{region 'Documentation'}
(*!
<summary>Restarts the scenario sequence and outer checks.</summary>
*)
{endregion}
METHOD PROTECTED ProcessReset
FScenario := ScenarioLowerLimits;
FChecked := FALSE;
FSubjectEnable := FALSE;
FEvaluateSubjects := FALSE;
FObservationReady := FALSE;
FFirstFailedScenario := 0;
FFailedDuringEvaluation := FALSE;
FCapture.Reset();
ResetSubjects();
FResults.Reset();
FActivity.Reset();
FInputs.Reset();
FFindings.Reset();
CompleteReset();
END_METHOD

{region 'Documentation'}
(*!
<summary>Consumes reset, evaluates, then waits for the outer checks before advancing.</summary>
*)
{endregion}
METHOD PROTECTED ProcessTests
VAR_INPUT
    Enable : BOOL; //! Phase permission supplied by the owning Test Case; FALSE does not authorize progression, while observation may continue.
END_VAR
IF NOT Enable THEN
    RETURN;
END_IF;

IF FChecked THEN
    FChecked := FALSE;
    FObservationReady := FALSE;
    IF FEvaluateSubjects THEN
        IF FScenario = LastScenario THEN
            CompleteTests();
            RETURN;
        END_IF;
        FScenario := FScenario + 1;
    END_IF;
    FEvaluateSubjects := NOT FEvaluateSubjects;
END_IF;

IF NOT SelectScenario() THEN
    RETURN;
END_IF;
FCapture.Reset();
IF NOT FEvaluateSubjects THEN
    ResetSubjects();
END_IF;

CallSubjects();
CheckResults();
CheckInputs();
CheckFindings();
IF (FFirstFailedScenario = 0)
    AND NOT (FResultsMatch AND FActivityMatch AND FInputsMatch AND FFindingsMatch) THEN
    FFirstFailedScenario := FScenario;
    FFailedDuringEvaluation := FEvaluateSubjects;
END_IF;
FObservationReady := TRUE;
END_METHOD

{region 'Documentation'}
(*!
<summary>Queues reset; the next bound FB call consumes it without evaluating.</summary>
*)
{endregion}
METHOD PRIVATE ResetSubjects
FSigned.Reset();
FUnsigned.Reset();
END_METHOD

{region 'Documentation'}
(*!
<summary>Selects explicit stimuli and expected results for one scenario.</summary>
*)
{endregion}
METHOD PRIVATE SelectScenario : BOOL //! TRUE after selecting a supported scenario and its literal expectations; FALSE reports an unknown scenario.
SelectScenario := FALSE;
FSubjectEnable := TRUE;
FSignedValue := -127;
FSignedMinimum := -128;
FUnsignedValue := 128;
FUnsignedMinimum := 128;
FUnsignedMaximum := 255;
CASE FScenario OF
    ScenarioLowerLimits:
        FSignedExpectedResult := E_Result.Passed;
        FSignedExpectedFinding := FALSE;
        FUnsignedExpectedResult := E_Result.Passed;
        FUnsignedExpectedFinding := FALSE;
    ScenarioUpperLimits:
        FSignedValue := 127;
        FUnsignedValue := 255;
        FSignedExpectedResult := E_Result.Passed;
        FSignedExpectedFinding := FALSE;
        FUnsignedExpectedResult := E_Result.Passed;
        FUnsignedExpectedFinding := FALSE;
    ScenarioEqualSignedMinimum:
        FSignedValue := -128;
        FSignedExpectedResult := E_Result.Failed;
        FSignedExpectedFinding := TRUE;
        FUnsignedExpectedResult := E_Result.Passed;
        FUnsignedExpectedFinding := FALSE;
    ScenarioOutsideRange:
        FSignedValue := -128;
        FSignedMinimum := -127;
        FUnsignedValue := 127;
        FSignedExpectedResult := E_Result.Failed;
        FSignedExpectedFinding := TRUE;
        FUnsignedExpectedResult := E_Result.Failed;
        FUnsignedExpectedFinding := TRUE;
    ScenarioAboveMaximum:
        FUnsignedValue := 255;
        FUnsignedMaximum := 254;
        FSignedExpectedResult := E_Result.Passed;
        FSignedExpectedFinding := FALSE;
        FUnsignedExpectedResult := E_Result.Failed;
        FUnsignedExpectedFinding := TRUE;
    ScenarioSingleValue:
        FUnsignedMinimum := 255;
        FUnsignedMaximum := 255;
        FUnsignedValue := 255;
        FSignedExpectedResult := E_Result.Passed;
        FSignedExpectedFinding := FALSE;
        FUnsignedExpectedResult := E_Result.Passed;
        FUnsignedExpectedFinding := FALSE;
    ScenarioReversedRange:
        FUnsignedMinimum := 255;
        FUnsignedMaximum := 128;
        FSignedExpectedResult := E_Result.Passed;
        FSignedExpectedFinding := FALSE;
        FUnsignedExpectedResult := E_Result.Error;
        FUnsignedExpectedFinding := TRUE;
ELSE
    Error(Message := 'Unknown variant Assertion scenario.');
    RETURN;
END_CASE;

SelectScenario := TRUE;
END_METHOD

END_FUNCTION_BLOCK

// ---- SelfTests/TestCases/TestSuite_AssertionVariants/Test_AssertionTemporalVariants.TcPOU
{region 'Documentation'}
(*!
<summary>Checks temporal variants with isolated production subjects.</summary>
<description>
Each independent scenario consumes a bound reset call before its evaluation call.
ProcessAssertions checks the observation before ProcessTests advances.
SelectScenario holds explicit expected results; no production algorithm is mirrored.
Expected findings remain in the local capture; only outer checks affect the test result.
FirstFailedScenario and FailedDuringEvaluation retain the first mismatch.
Each scenario uses literal typed inputs at the declared operand widths.
</description>
*)
{endregion}
FUNCTION_BLOCK Test_AssertionTemporalVariants EXTENDS TestCaseBase
VAR
    FTimestamp : AssertEqual_LDT;
    FTimestampExpectedResult : E_Result;
    FTimestampExpectedFinding : BOOL;
    FTimespan : AssertInTimespan_DT;
    FTimespanExpectedResult : E_Result;
    FTimespanExpectedFinding : BOOL;

    FTimestampValue : LDT;
    FExpectedTimestamp : LDT;
    FTime : DT;
    FStartTime : DT;
    FEndTime : DT;
    FSubjectEnable : BOOL;
    FCapture : EventBuffer;
    FEvents : ARRAY[1..CaptureLength] OF ST_Event;
    FCaptureFifo : ST_FifoStatus;
    FCaptureStatus : ST_EventBufferStatus;
    FSetupValid : BOOL;
    FScenario : UINT;
    FChecked : BOOL;
    FEvaluateSubjects : BOOL;
    FObservationReady : BOOL;
    FFirstFailedScenario : UINT;
    FFailedDuringEvaluation : BOOL;
    FResultsMatch : BOOL;
    FResults : AssertTrue;
    FActivityMatch : BOOL;
    FActivity : AssertTrue;
    FInputsMatch : BOOL;
    FInputs : AssertTrue;
    FFindingsMatch : BOOL;
    FFindings : AssertTrue;
END_VAR
VAR CONSTANT
    CaptureLength : UINT := 8;
    ScenarioLowerBound : UINT := 1;
    ScenarioUpperBound : UINT := 2;
    ScenarioNanosecondDifference : UINT := 3;
    ScenarioBeforeStart : UINT := 4;
    ScenarioAfterEnd : UINT := 5;
    ScenarioSingleInstant : UINT := 6;
    ScenarioReversedTimespan : UINT := 7;
    LastScenario : UINT := ScenarioReversedTimespan;
END_VAR

SUPER^();

{region 'Documentation'}
(*!
<summary>Aggregates only outer checks, not intentionally failing subjects.</summary>
*)
{endregion}
METHOD PROTECTED AggregateResults
VAR_INPUT
    Aggregator : I_ResultAggregator; //! Borrowed result sink owned by the outer Test Case; add this test's checking Assertions without resetting or retaining the sink.
END_VAR
Aggregator.AddProvider(Provider := FResults);
Aggregator.AddProvider(Provider := FActivity);
Aggregator.AddProvider(Provider := FInputs);
Aggregator.AddProvider(Provider := FFindings);
END_METHOD

{region 'Documentation'}
(*!
<summary>Calls each inherited production subject once with caller-owned input storage.</summary>
*)
{endregion}
METHOD PRIVATE CallSubjects
FTimestamp(Enable := FSubjectEnable,
    State := E_State.Running,
    IN := FTimestampValue,
    Expected := FExpectedTimestamp);
FTimespan(Enable := FSubjectEnable,
    State := E_State.Running,
    IN := FTime,
    StartTime := FStartTime,
    EndTime := FEndTime);
END_METHOD

{region 'Documentation'}
(*!
<summary>Checks one subject finding in call order; expected outcomes come from the scenario.</summary>
*)
{endregion}
METHOD PRIVATE CheckFinding : BOOL //! TRUE when the required finding checks pass; calls requiring no finding also succeed.
VAR_INPUT
    Subject : I_Assertion; //! Assertion interface supplying the expected finding identity.
    ExpectedResult : E_Result; //! Independently authored result expected in the captured finding.
    ExpectedFinding : BOOL; //! TRUE when this scenario requires a finding during active evaluation.
END_VAR
VAR_IN_OUT
    Index : UINT; //! One-based next finding index; advanced when this call checks a required finding.
END_VAR
CheckFinding := TRUE;
IF FEvaluateSubjects AND ExpectedFinding THEN
    CheckFinding := (FEvents[Index].SequenceId = UINT_TO_UDINT(Index))
        AND (FEvents[Index].Name = Subject.Name)
        AND (FEvents[Index].OwnerScope = E_OwnerScope.Assertion)
        AND (FEvents[Index].EventType = E_EventType.Result)
        AND (FEvents[Index].State = E_State.Running)
        AND (FEvents[Index].Result = ExpectedResult)
        AND (FEvents[Index].Message <> '');
    Index := Index + 1;
END_IF;
END_METHOD

{region 'Documentation'}
(*!
<summary>Checks exact finding count and identities; at most one finding per subject.</summary>
*)
{endregion}
METHOD PRIVATE CheckFindings
VAR
    Index : UINT;
    Matches : BOOL;
END_VAR
Index := 1;
FFindingsMatch := TRUE;
Matches := CheckFinding(Subject := FTimestamp,
    ExpectedResult := FTimestampExpectedResult,
    ExpectedFinding := FTimestampExpectedFinding,
    Index := Index);
FFindingsMatch := FFindingsMatch AND Matches;
Matches := CheckFinding(Subject := FTimespan,
    ExpectedResult := FTimespanExpectedResult,
    ExpectedFinding := FTimespanExpectedFinding,
    Index := Index);
FFindingsMatch := FFindingsMatch AND Matches;
FFindingsMatch := FFindingsMatch
    AND (FCaptureStatus.SequenceId = UINT_TO_UDINT(Index - 1))
    AND (FCaptureStatus.LostEventCount = 0);
END_METHOD

{region 'Documentation'}
(*!
<summary>Rejects incomplete subject, capture or outer Assertion setup.</summary>
*)
{endregion}
METHOD PROTECTED CheckInitialization : BOOL //! TRUE when the inherited initialization check and this concrete fixture check both accept the setup.
CheckInitialization := SUPER^.CheckInitialization();
IF NOT CheckInitialization THEN
    RETURN;
END_IF;

CheckInitialization := FSetupValid
    AND FResults.IsInitialized
    AND FActivity.IsInitialized
    AND FInputs.IsInitialized
    AND FFindings.IsInitialized;
IF NOT CheckInitialization THEN
    EventPublisher.PublishEvent(Event := CreateFrameworkEvent(Name := Name,
        ResourceName := '',
        State := State,
        Severity := E_EventSeverity.Error,
        Message := 'Variant selftest setup failed.'));
END_IF;
END_METHOD

{region 'Documentation'}
(*!
<summary>Verifies input preservation without using the tested comparison algorithm.</summary>
*)
{endregion}
METHOD PRIVATE CheckInputs
FInputsMatch := (FTimestamp.IN = FTimestampValue)
    AND (FTimestamp.Expected = FExpectedTimestamp)
    AND (FTimespan.IN = FTime)
    AND (FTimespan.StartTime = FStartTime)
    AND (FTimespan.EndTime = FEndTime);
END_METHOD

{region 'Documentation'}
(*!
<summary>Checks literal evaluation results, or NotEvaluated on the reset call.</summary>
*)
{endregion}
METHOD PRIVATE CheckResults
IF FEvaluateSubjects THEN
    FResultsMatch := (FTimestamp.Result = FTimestampExpectedResult)
        AND (FTimespan.Result = FTimespanExpectedResult);
ELSE
    FResultsMatch := (FTimestamp.Result = E_Result.NotEvaluated)
        AND (FTimespan.Result = E_Result.NotEvaluated);
END_IF;
FActivityMatch := (FTimestamp.Enabled = FSubjectEnable)
    AND (FTimestamp.ObservationActive = (FEvaluateSubjects AND FSubjectEnable))
    AND (FTimestamp.EvaluationActive = (FEvaluateSubjects AND FSubjectEnable))
    AND (FTimespan.Enabled = FSubjectEnable)
    AND (FTimespan.ObservationActive = (FEvaluateSubjects AND FSubjectEnable))
    AND (FTimespan.EvaluationActive = (FEvaluateSubjects AND FSubjectEnable));
END_METHOD

{region 'Documentation'}
(*!
<summary>Initializes outer checks and isolates intentional subject findings.</summary>
*)
{endregion}
METHOD PROTECTED Configure
VAR
    Initialized : BOOL;
END_VAR
FPreparationStateCount := 0;
FTestStateCount := 1;
FResults.Initialize(Parent := THIS^,
    AssertionName := 'Results');
FActivity.Initialize(Parent := THIS^,
    AssertionName := 'Activity');
FInputs.Initialize(Parent := THIS^,
    AssertionName := 'Inputs');
FFindings.Initialize(Parent := THIS^,
    AssertionName := 'Findings');
FSetupValid := FCapture.Initialize(Buffer := FEvents,
    FifoControl := FCaptureFifo,
    Status := FCaptureStatus);
FTimestamp.BindPublisher(Publisher := FCapture);
Initialized := FTimestamp.Initialize(Parent := THIS^,
    AssertionName := 'Timestamp');
FSetupValid := FSetupValid AND Initialized;
FTimespan.BindPublisher(Publisher := FCapture);
Initialized := FTimespan.Initialize(Parent := THIS^,
    AssertionName := 'Timespan');
FSetupValid := FSetupValid AND Initialized;
END_METHOD

{region 'Documentation'}
(*!
<summary>Completes abort; no asynchronous resource is owned.</summary>
*)
{endregion}
METHOD PROTECTED ProcessAbort
VAR_INPUT
    Enable : BOOL; //! Phase permission supplied by the owning Test Case; FALSE does not authorize progression, while observation may continue.
END_VAR
IF Enable THEN
    CompleteAbort();
END_IF;
END_METHOD

{region 'Documentation'}
(*!
<summary>Latches this call's checks before progression is permitted.</summary>
*)
{endregion}
METHOD PROTECTED ProcessAssertions
VAR_INPUT
    Enable : BOOL; //! Phase permission supplied by the owning Test Case; FALSE does not authorize progression, while observation may continue.
END_VAR
VAR
    Check : BOOL;
END_VAR
Check := Enable AND FObservationReady;
FResults(Enable := Check,
    State := State,
    IN := FResultsMatch);
FActivity(Enable := Check,
    State := State,
    IN := FActivityMatch);
FInputs(Enable := Check,
    State := State,
    IN := FInputsMatch);
FFindings(Enable := Check,
    State := State,
    IN := FFindingsMatch);
IF Check THEN
    FChecked := TRUE;
END_IF;
END_METHOD

{region 'Documentation'}
(*!
<summary>No Preparation phase is needed.</summary>
*)
{endregion}
METHOD PROTECTED ProcessPreparations
VAR_INPUT
    // SA0033: Required hook; this test has no Preparation phase.
    {attribute 'analysis' := '-33'}
    Enable : BOOL; //! Phase permission supplied by the owning Test Case; FALSE does not authorize progression, while observation may continue.
END_VAR
END_METHOD

{region 'Documentation'}
(*!
<summary>Restarts the scenario sequence and outer checks.</summary>
*)
{endregion}
METHOD PROTECTED ProcessReset
FScenario := ScenarioLowerBound;
FChecked := FALSE;
FSubjectEnable := FALSE;
FEvaluateSubjects := FALSE;
FObservationReady := FALSE;
FFirstFailedScenario := 0;
FFailedDuringEvaluation := FALSE;
FCapture.Reset();
ResetSubjects();
FResults.Reset();
FActivity.Reset();
FInputs.Reset();
FFindings.Reset();
CompleteReset();
END_METHOD

{region 'Documentation'}
(*!
<summary>Consumes reset, evaluates, then waits for the outer checks before advancing.</summary>
*)
{endregion}
METHOD PROTECTED ProcessTests
VAR_INPUT
    Enable : BOOL; //! Phase permission supplied by the owning Test Case; FALSE does not authorize progression, while observation may continue.
END_VAR
IF NOT Enable THEN
    RETURN;
END_IF;

IF FChecked THEN
    FChecked := FALSE;
    FObservationReady := FALSE;
    IF FEvaluateSubjects THEN
        IF FScenario = LastScenario THEN
            CompleteTests();
            RETURN;
        END_IF;
        FScenario := FScenario + 1;
    END_IF;
    FEvaluateSubjects := NOT FEvaluateSubjects;
END_IF;

IF NOT SelectScenario() THEN
    RETURN;
END_IF;
FCapture.Reset();
IF NOT FEvaluateSubjects THEN
    ResetSubjects();
END_IF;

CallSubjects();
CheckResults();
CheckInputs();
CheckFindings();
IF (FFirstFailedScenario = 0)
    AND NOT (FResultsMatch AND FActivityMatch AND FInputsMatch AND FFindingsMatch) THEN
    FFirstFailedScenario := FScenario;
    FFailedDuringEvaluation := FEvaluateSubjects;
END_IF;
FObservationReady := TRUE;
END_METHOD

{region 'Documentation'}
(*!
<summary>Queues reset; the next bound FB call consumes it without evaluating.</summary>
*)
{endregion}
METHOD PRIVATE ResetSubjects
FTimestamp.Reset();
FTimespan.Reset();
END_METHOD

{region 'Documentation'}
(*!
<summary>Selects explicit stimuli and expected results for one scenario.</summary>
*)
{endregion}
METHOD PRIVATE SelectScenario : BOOL //! TRUE after selecting a supported scenario and its literal expectations; FALSE reports an unknown scenario.
SelectScenario := FALSE;
FSubjectEnable := TRUE;
FTimestampValue := LDT#2026-01-02-03:04:05.000000001;
FExpectedTimestamp := LDT#2026-01-02-03:04:05.000000001;
FTime := DT#2026-01-02-03:04:05;
FStartTime := DT#2026-01-02-03:04:05;
FEndTime := DT#2026-01-02-03:04:07;
CASE FScenario OF
    ScenarioLowerBound:
        FTimestampExpectedResult := E_Result.Passed;
        FTimestampExpectedFinding := FALSE;
        FTimespanExpectedResult := E_Result.Passed;
        FTimespanExpectedFinding := FALSE;
    ScenarioUpperBound:
        FTime := DT#2026-01-02-03:04:07;
        FTimestampExpectedResult := E_Result.Passed;
        FTimestampExpectedFinding := FALSE;
        FTimespanExpectedResult := E_Result.Passed;
        FTimespanExpectedFinding := FALSE;
    ScenarioNanosecondDifference:
        FTimestampValue := LDT#2026-01-02-03:04:05.000000002;
        FTimestampExpectedResult := E_Result.Failed;
        FTimestampExpectedFinding := TRUE;
        FTimespanExpectedResult := E_Result.Passed;
        FTimespanExpectedFinding := FALSE;
    ScenarioBeforeStart:
        FTime := DT#2026-01-02-03:04:04;
        FTimestampExpectedResult := E_Result.Passed;
        FTimestampExpectedFinding := FALSE;
        FTimespanExpectedResult := E_Result.Failed;
        FTimespanExpectedFinding := TRUE;
    ScenarioAfterEnd:
        FTime := DT#2026-01-02-03:04:08;
        FTimestampExpectedResult := E_Result.Passed;
        FTimestampExpectedFinding := FALSE;
        FTimespanExpectedResult := E_Result.Failed;
        FTimespanExpectedFinding := TRUE;
    ScenarioSingleInstant:
        FEndTime := FStartTime;
        FTimestampExpectedResult := E_Result.Passed;
        FTimestampExpectedFinding := FALSE;
        FTimespanExpectedResult := E_Result.Passed;
        FTimespanExpectedFinding := FALSE;
    ScenarioReversedTimespan:
        FStartTime := DT#2026-01-02-03:04:07;
        FEndTime := DT#2026-01-02-03:04:05;
        FTimestampExpectedResult := E_Result.Passed;
        FTimestampExpectedFinding := FALSE;
        FTimespanExpectedResult := E_Result.Error;
        FTimespanExpectedFinding := TRUE;
ELSE
    Error(Message := 'Unknown variant Assertion scenario.');
    RETURN;
END_CASE;

SelectScenario := TRUE;
END_METHOD

END_FUNCTION_BLOCK

// ---- Framework/Assertions/POU/BasicTypes/LDT/AssertEqual_LDT.TcPOU
{region 'Documentation'}
(*!
<summary>Checks equality with the expected LDT value.</summary>
*)
{endregion}
FUNCTION_BLOCK AssertEqual_LDT EXTENDS AssertionBase
VAR_INPUT
    IN : LDT; //! Actual value checked or observed by this Assertion.
    Expected : LDT; //! Reference value for comparison with IN.
END_VAR

SUPER^();

{region 'Documentation'}
(*!
<summary>Evaluate the typed temporal relation and report higher-priority errors first.</summary>
*)
{endregion}
METHOD PROTECTED Assert
VAR
    Message : STRING(GVL_Constants.MessageLength);
    ExpectedText : STRING(GVL_Constants.AssertionValueLength);
    ActualText : STRING(GVL_Constants.AssertionValueLength);
END_VAR
IF NOT EvaluationActive THEN
    RETURN;
END_IF;

IF Result = E_Result.Error THEN
    RETURN;
END_IF;

IF Result = E_Result.Failed THEN
    RETURN;
END_IF;

IF IN <> Expected THEN
    ExpectedText := LDT_TO_STRING(Expected);
    ActualText := LDT_TO_STRING(IN);
    Message := CONCAT('Assertion failed: values are not equal. Expected = ',
        ExpectedText);
    Message := CONCAT(Message, ', Actual = ');
    Message := CONCAT(Message, ActualText);
    Message := CONCAT(Message, '.');
    Fail(Message := Message);
    RETURN;
END_IF;

Pass();
END_METHOD

END_FUNCTION_BLOCK

// ---- Framework/Assertions/POU/BasicTypes/DT/AssertInTimespan_DT.TcPOU
{region 'Documentation'}
(*!
<summary>Check that IN is inside the inclusive StartTime..EndTime interval.</summary>
<description>

StartTime &gt; EndTime reports Error during active evaluation; equal bounds are
valid.

</description>
*)
{endregion}
FUNCTION_BLOCK AssertInTimespan_DT EXTENDS AssertionBase
VAR_INPUT
    IN : DT; //! Actual value checked or observed by this Assertion.
    StartTime : DT; //! Inclusive start of the time span; must not exceed EndTime.
    EndTime : DT; //! Inclusive end of the time span; must not precede StartTime.
END_VAR

SUPER^();

{region 'Documentation'}
(*!
<summary>Evaluate the typed temporal relation and report higher-priority errors first.</summary>
*)
{endregion}
METHOD PROTECTED Assert
VAR
    Message : STRING(GVL_Constants.MessageLength);
    StartTimeText : STRING(GVL_Constants.AssertionValueLength);
    EndTimeText : STRING(GVL_Constants.AssertionValueLength);
    ActualText : STRING(GVL_Constants.AssertionValueLength);
END_VAR
IF NOT EvaluationActive THEN
    RETURN;
END_IF;

IF Result = E_Result.Error THEN
    RETURN;
END_IF;

IF StartTime > EndTime THEN
    StartTimeText := DT_TO_STRING(StartTime);
    EndTimeText := DT_TO_STRING(EndTime);
    Message := CONCAT('Assertion error: start time exceeds end time. StartTime = ',
        StartTimeText);
    Message := CONCAT(Message, ', EndTime = ');
    Message := CONCAT(Message, EndTimeText);
    Message := CONCAT(Message, '.');
    Error(Message := Message);
    RETURN;
END_IF;

IF Result = E_Result.Failed THEN
    RETURN;
END_IF;

IF (IN < StartTime) OR (IN > EndTime) THEN
    StartTimeText := DT_TO_STRING(StartTime);
    EndTimeText := DT_TO_STRING(EndTime);
    ActualText := DT_TO_STRING(IN);
    Message := CONCAT('Assertion failed: value is outside allowed timespan. StartTime = ',
        StartTimeText);
    Message := CONCAT(Message, ', EndTime = ');
    Message := CONCAT(Message, EndTimeText);
    Message := CONCAT(Message, ', Actual = ');
    Message := CONCAT(Message, ActualText);
    Message := CONCAT(Message, '.');
    Fail(Message := Message);
    RETURN;
END_IF;

Pass();
END_METHOD

END_FUNCTION_BLOCK

// ---- Framework/Common/POU/GetFrameworkVersion.TcPOU
{region 'Documentation'}
(*!
<summary>Returns Major.Minor.Build from the generated library metadata; revision is omitted.</summary>
*)
{endregion}
FUNCTION GetFrameworkVersion : STRING(GVL_Constants.VersionLength) //! Library version as Major.Minor.Build without revision, within VersionLength.

GetFrameworkVersion := UINT_TO_STRING(Global_Version.stLibVersion_Tc3_UnitTest.iMajor);
GetFrameworkVersion := CONCAT(GetFrameworkVersion, '.');
GetFrameworkVersion := CONCAT(GetFrameworkVersion, UINT_TO_STRING(Global_Version.stLibVersion_Tc3_UnitTest.iMinor));
GetFrameworkVersion := CONCAT(GetFrameworkVersion, '.');
GetFrameworkVersion := CONCAT(GetFrameworkVersion, UINT_TO_STRING(Global_Version.stLibVersion_Tc3_UnitTest.iBuild));

END_FUNCTION

// ---- Framework/Assertions/POU/Arrays/Bool/AssertArrayContainsArray_Bool.TcPOU
{region 'Documentation'}
(*!
<summary>Searches the selected IN range for the complete contiguous Expected pattern.</summary>
<description>

StartIndex is an absolute declared IN index, not an offset. Length selects 1..255
elements; the complete selected range must fit IN. Invalid references or ranges report
Error.

Keep supplied arrays stable for the call. Input data is read, not copied or retained as a
snapshot.

The complete Expected pattern must be nonempty and fit the selected IN range; an
oversized pattern reports Error, not a missing-match result.

</description>
*)
{endregion}
FUNCTION_BLOCK AssertArrayContainsArray_Bool EXTENDS AssertionBase
VAR_INPUT
    StartIndex : DINT; //! First selected index in IN; uses the array's declared index range, not a zero-based offset.
    Length : USINT; //! Number of searched elements, from 1 through 255.
END_VAR
VAR_IN_OUT CONSTANT
    IN : ARRAY[*] OF BOOL; //! Read-only search data; keep stable during the call.
    Expected : ARRAY[*] OF BOOL; //! Read-only expected sequence starting at its own lower bound; must fit the selected actual range.
END_VAR

SUPER^();

{region 'Documentation'}
(*!
<summary>Validate configuration before searching the selected range.</summary>
*)
{endregion}
METHOD PROTECTED Assert
VAR
    InLowerIndex : DINT;
    InUpperIndex : DINT;
    EndIndex : LINT;
    Offset : LINT;
    InIndex : DINT;
    ExpectedLowerIndex : DINT;
    ExpectedUpperIndex : DINT;
    ExpectedLength : LINT;
    ExpectedIndex : DINT;
    CandidateOffset : LINT;
    PatternFound : BOOL;
    PatternMatches : BOOL;
    Message : STRING(GVL_Constants.MessageLength);
END_VAR
IF NOT EvaluationActive THEN
    RETURN;
END_IF;

IF Result = E_Result.Error THEN
    RETURN;
END_IF;

// C0371: FB input is checked here before any reference access.
{warning disable C0371}
IF NOT __ISVALIDREF(IN) THEN
    Error(Message := 'Assertion error: IN reference is invalid.');
    RETURN;
END_IF;

IF NOT __ISVALIDREF(Expected) THEN
    Error(Message := 'Assertion error: Expected reference is invalid.');
    RETURN;
END_IF;

InLowerIndex := LOWER_BOUND(IN, 1);
InUpperIndex := UPPER_BOUND(IN, 1);
EndIndex := DINT_TO_LINT(StartIndex) + USINT_TO_LINT(Length) - 1;

ExpectedLowerIndex := LOWER_BOUND(Expected, 1);
ExpectedUpperIndex := UPPER_BOUND(Expected, 1);
ExpectedLength := DINT_TO_LINT(ExpectedUpperIndex) - DINT_TO_LINT(ExpectedLowerIndex) + 1;

IF (Length = 0)
    OR (ExpectedLength <= 0) OR (ExpectedLength > USINT_TO_LINT(Length))
    OR (StartIndex < InLowerIndex) OR (StartIndex > InUpperIndex)
    OR (EndIndex > DINT_TO_LINT(InUpperIndex)) THEN
    Message := CONCAT('Assertion error: array range or pattern is invalid. StartIndex = ',
        DINT_TO_STRING(StartIndex));
    Message := CONCAT(Message, ', Length = ');
    Message := CONCAT(Message, USINT_TO_STRING(Length));
    Message := CONCAT(Message, ', ExpectedLength = ');
    Message := CONCAT(Message, LINT_TO_STRING(ExpectedLength));
    Message := CONCAT(Message, '.');
    Error(Message := Message);
    RETURN;
END_IF;

IF Result = E_Result.Failed THEN
    RETURN;
END_IF;

PatternFound := FALSE;
FOR CandidateOffset := 0 TO USINT_TO_LINT(Length) - ExpectedLength DO
    PatternMatches := TRUE;
    FOR Offset := 0 TO ExpectedLength - 1 DO
        InIndex := LINT_TO_DINT(DINT_TO_LINT(StartIndex) + CandidateOffset + Offset);
        ExpectedIndex := LINT_TO_DINT(DINT_TO_LINT(ExpectedLowerIndex) + Offset);
        IF IN[InIndex] <> Expected[ExpectedIndex] THEN
            PatternMatches := FALSE;
            EXIT;
        END_IF;
    END_FOR;

    IF PatternMatches THEN
        PatternFound := TRUE;
        EXIT;
    END_IF;
END_FOR;

IF NOT PatternFound THEN
    Message := CONCAT('Assertion failed: array range does not contain Expected pattern. ExpectedRange = [',
        DINT_TO_STRING(ExpectedLowerIndex));
    Message := CONCAT(Message, '..');
    Message := CONCAT(Message, DINT_TO_STRING(ExpectedUpperIndex));
    Message := CONCAT(Message, '], ActualRange = [');
    Message := CONCAT(Message, DINT_TO_STRING(StartIndex));
    Message := CONCAT(Message, '..');
    Message := CONCAT(Message, LINT_TO_STRING(EndIndex));
    Message := CONCAT(Message, ']');
    Message := CONCAT(Message, '.');
    Fail(Message := Message);
    RETURN;
END_IF;

Pass();
{warning restore C0371}
END_METHOD

END_FUNCTION_BLOCK

// ---- Framework/Assertions/POU/Arrays/Bool/AssertArrayNoValueChange_Bool.TcPOU
{region 'Documentation'}
(*!
<summary>Captures one snapshot until Reset; Disable/Re-Enable never replaces it.</summary>
<description>

Disabling observation preserves the original snapshot. Re-enabling requires a fresh
preceding observation before comparisons resume; it does not replace that snapshot.

StartIndex is an absolute IN index and Length selects 1..255 elements within IN. Memory
must have at least Length elements from its own lower bound. Invalid references or ranges
report Error.

The caller provides dedicated writable Memory that must not overlap IN; overlap is not
checked. Keep bindings, selected range and snapshot contents stable until Reset. Reset
invalidates the snapshot without clearing Memory bytes.

</description>
*)
{endregion}
FUNCTION_BLOCK AssertArrayNoValueChange_Bool EXTENDS AssertionBase
VAR_INPUT
    StartIndex : DINT; //! First selected index in IN; uses the array's declared index range, not a zero-based offset.
    Length : USINT; //! Number of monitored elements, from 1 through 255.
END_VAR
VAR_IN_OUT CONSTANT
    IN : ARRAY[*] OF BOOL; //! Read-only actual data; the selected range must remain stable during the call.
END_VAR
VAR_IN_OUT
    Memory : ARRAY[*] OF BOOL; //! Dedicated snapshot storage; only this assertion writes its selected elements.
END_VAR
VAR
    FSnapshotValid : BOOL;
    FObservationPrevious : BOOL;
    FEvaluationActive : BOOL;
END_VAR

SUPER^();

{region 'Documentation'}
(*!
<summary>Capture once or compare against the retained snapshot after range validation.</summary>
*)
{endregion}
METHOD PROTECTED Assert
VAR
    InLowerIndex : DINT;
    InUpperIndex : DINT;
    MemoryLowerIndex : DINT;
    MemoryUpperIndex : DINT;
    MemoryEndIndex : LINT;
    EndIndex : LINT;
    Offset : LINT;
    InIndex : DINT;
    MemoryIndex : DINT;
    Message : STRING(GVL_Constants.MessageLength);
    ReferenceText : STRING(GVL_Constants.AssertionValueLength);
    ActualText : STRING(GVL_Constants.AssertionValueLength);
END_VAR
FEvaluationActive := ObservationActive AND FObservationPrevious AND FSnapshotValid;
FObservationPrevious := ObservationActive;

IF NOT ObservationActive THEN
    RETURN;
END_IF;

IF Result = E_Result.Error THEN
    RETURN;
END_IF;

// C0371: FB inputs are checked here before any reference access.
{warning disable C0371}
IF NOT __ISVALIDREF(IN) THEN
    Error(Message := 'Assertion error: IN reference is invalid.');
    RETURN;
END_IF;

IF NOT __ISVALIDREF(Memory) THEN
    Error(Message := 'Assertion error: Memory reference is invalid.');
    RETURN;
END_IF;

InLowerIndex := LOWER_BOUND(IN, 1);
InUpperIndex := UPPER_BOUND(IN, 1);
MemoryLowerIndex := LOWER_BOUND(Memory, 1);
MemoryUpperIndex := UPPER_BOUND(Memory, 1);
EndIndex := DINT_TO_LINT(StartIndex) + USINT_TO_LINT(Length) - 1;
MemoryEndIndex := DINT_TO_LINT(MemoryLowerIndex) + USINT_TO_LINT(Length) - 1;

IF (Length = 0)
    OR (StartIndex < InLowerIndex) OR (StartIndex > InUpperIndex)
    OR (EndIndex > DINT_TO_LINT(InUpperIndex))
    OR (MemoryEndIndex > DINT_TO_LINT(MemoryUpperIndex)) THEN
    Message := CONCAT('Assertion error: array or memory range is invalid. StartIndex = ',
        DINT_TO_STRING(StartIndex));
    Message := CONCAT(Message, ', EndIndex = ');
    Message := CONCAT(Message, LINT_TO_STRING(EndIndex));
    Message := CONCAT(Message, ', Length = ');
    Message := CONCAT(Message, USINT_TO_STRING(Length));
    Message := CONCAT(Message, '.');
    Error(Message := Message);
    RETURN;
END_IF;

IF NOT FSnapshotValid THEN
    FOR Offset := 0 TO USINT_TO_LINT(Length) - 1 DO
        InIndex := LINT_TO_DINT(DINT_TO_LINT(StartIndex) + Offset);
        MemoryIndex := LINT_TO_DINT(DINT_TO_LINT(MemoryLowerIndex) + Offset);
        Memory[MemoryIndex] := IN[InIndex];
    END_FOR;
    FSnapshotValid := TRUE;
    RETURN;
END_IF;

IF NOT EvaluationActive THEN
    RETURN;
END_IF;

IF Result = E_Result.Failed THEN
    RETURN;
END_IF;

FOR Offset := 0 TO USINT_TO_LINT(Length) - 1 DO
    InIndex := LINT_TO_DINT(DINT_TO_LINT(StartIndex) + Offset);
    MemoryIndex := LINT_TO_DINT(DINT_TO_LINT(MemoryLowerIndex) + Offset);
    IF IN[InIndex] <> Memory[MemoryIndex] THEN
        ReferenceText := BOOL_TO_STRING(Memory[MemoryIndex]);
        ActualText := BOOL_TO_STRING(IN[InIndex]);
        Message := CONCAT('Assertion failed: array value changed. Reference[',
            DINT_TO_STRING(MemoryIndex));
        Message := CONCAT(Message, '] = ');
        Message := CONCAT(Message, ReferenceText);
        Message := CONCAT(Message, ', IN[');
        Message := CONCAT(Message, DINT_TO_STRING(InIndex));
        Message := CONCAT(Message, '] = ');
        Message := CONCAT(Message, ActualText);
        Message := CONCAT(Message, '.');
        Fail(Message := Message);
        RETURN;
    END_IF;
END_FOR;

Pass();
{warning restore C0371}
END_METHOD

{region 'Documentation'}
(*!
<summary>Current/last call has consecutive observation and an existing snapshot.</summary>
*)
{endregion}
{attribute 'monitoring' := 'call'}
PROPERTY PUBLIC EvaluationActive : BOOL //! Current/last call has consecutive observation and an existing snapshot.
GET // PUBLIC
EvaluationActive := FEvaluationActive;
END_GET
END_PROPERTY

{region 'Documentation'}
(*!
<summary>Invalidate the snapshot and observation history.</summary>
<description>

Does not clear external Memory. The next active observation captures a new snapshot
before comparison.

</description>
*)
{endregion}
METHOD PROTECTED ResetAssertion
FSnapshotValid := FALSE;
FObservationPrevious := FALSE;
FEvaluationActive := FALSE;
END_METHOD

END_FUNCTION_BLOCK

// ---- Framework/Assertions/POU/Arrays/Bool/AssertEqualArray_Bool.TcPOU
{region 'Documentation'}
(*!
<summary>Compares the entire Expected array with IN starting at StartIndex.</summary>
<description>

StartIndex is an absolute declared IN index. The entire Expected array, starting at its
own lower bound, determines the compared length and must fit IN. Invalid references or ranges
report Error.

Keep supplied arrays stable for the call. Input data is read, not copied or retained as a
snapshot.

</description>
*)
{endregion}
FUNCTION_BLOCK AssertEqualArray_Bool EXTENDS AssertionBase
VAR_INPUT
    StartIndex : DINT; //! First compared index in IN; Expected starts at its own lower bound.
END_VAR
VAR_IN_OUT CONSTANT
    IN : ARRAY[*] OF BOOL; //! Read-only actual data; the selected range must remain stable during the call.
    Expected : ARRAY[*] OF BOOL; //! Read-only expected sequence starting at its own lower bound; must fit the selected actual range.
END_VAR

SUPER^();

{region 'Documentation'}
(*!
<summary>Validate the selected range and expectations before comparing elements.</summary>
*)
{endregion}
METHOD PROTECTED Assert
VAR
    InLowerIndex : DINT;
    InUpperIndex : DINT;
    ExpectedLowerIndex : DINT;
    ExpectedUpperIndex : DINT;
    ExpectedLength : LINT;
    EndIndex : LINT;
    Offset : LINT;
    InIndex : DINT;
    ExpectedIndex : DINT;
    Message : STRING(GVL_Constants.MessageLength);
    ExpectedText : STRING(GVL_Constants.AssertionValueLength);
    ActualText : STRING(GVL_Constants.AssertionValueLength);
END_VAR
IF NOT EvaluationActive THEN
    RETURN;
END_IF;

IF Result = E_Result.Error THEN
    RETURN;
END_IF;

// C0371: FB inputs are checked here before any reference access.
{warning disable C0371}
IF NOT __ISVALIDREF(IN) THEN
    Error(Message := 'Assertion error: IN reference is invalid.');
    RETURN;
END_IF;

IF NOT __ISVALIDREF(Expected) THEN
    Error(Message := 'Assertion error: Expected reference is invalid.');
    RETURN;
END_IF;

InLowerIndex := LOWER_BOUND(IN, 1);
InUpperIndex := UPPER_BOUND(IN, 1);
ExpectedLowerIndex := LOWER_BOUND(Expected, 1);
ExpectedUpperIndex := UPPER_BOUND(Expected, 1);
ExpectedLength := DINT_TO_LINT(ExpectedUpperIndex) - DINT_TO_LINT(ExpectedLowerIndex) + 1;
EndIndex := DINT_TO_LINT(StartIndex) + ExpectedLength - 1;

IF (ExpectedLength <= 0)
    OR (StartIndex < InLowerIndex) OR (StartIndex > InUpperIndex)
    OR (EndIndex > DINT_TO_LINT(InUpperIndex)) THEN
    Message := CONCAT('Assertion error: array range is invalid. StartIndex = ',
        DINT_TO_STRING(StartIndex));
    Message := CONCAT(Message, ', EndIndex = ');
    Message := CONCAT(Message, LINT_TO_STRING(EndIndex));
    Message := CONCAT(Message, ', InLowerIndex = ');
    Message := CONCAT(Message, DINT_TO_STRING(InLowerIndex));
    Message := CONCAT(Message, ', InUpperIndex = ');
    Message := CONCAT(Message, DINT_TO_STRING(InUpperIndex));
    Message := CONCAT(Message, ', ExpectedLength = ');
    Message := CONCAT(Message, LINT_TO_STRING(ExpectedLength));
    Message := CONCAT(Message, '.');
    Error(Message := Message);
    RETURN;
END_IF;

IF Result = E_Result.Failed THEN
    RETURN;
END_IF;

FOR Offset := 0 TO ExpectedLength - 1 DO
    InIndex := LINT_TO_DINT(DINT_TO_LINT(StartIndex) + Offset);
    ExpectedIndex := LINT_TO_DINT(DINT_TO_LINT(ExpectedLowerIndex) + Offset);
    IF IN[InIndex] <> Expected[ExpectedIndex] THEN
        ExpectedText := BOOL_TO_STRING(Expected[ExpectedIndex]);
        ActualText := BOOL_TO_STRING(IN[InIndex]);
        Message := CONCAT('Assertion failed: array elements differ. Expected[',
            DINT_TO_STRING(ExpectedIndex));
        Message := CONCAT(Message, '] = ');
        Message := CONCAT(Message, ExpectedText);
        Message := CONCAT(Message, ', IN[');
        Message := CONCAT(Message, DINT_TO_STRING(InIndex));
        Message := CONCAT(Message, '] = ');
        Message := CONCAT(Message, ActualText);
        Message := CONCAT(Message, '.');
        Fail(Message := Message);
        RETURN;
    END_IF;
END_FOR;

Pass();
{warning restore C0371}
END_METHOD

END_FUNCTION_BLOCK

// ---- Framework/Assertions/POU/Arrays/Byte/AssertArrayAllEqual_Byte.TcPOU
{region 'Documentation'}
(*!
<summary>Checks every selected IN element against Expected; reports the first
mismatch.</summary>
<description>

StartIndex is an absolute declared IN index, not an offset. Length selects 1..255
elements; the complete selected range must fit IN. Invalid references or ranges report
Error.

Keep supplied arrays stable for the call. Input data is read, not copied or retained as a
snapshot.

Comparison applies Mask to both values; bits outside it are ignored. The default mask
selects all bits.

</description>
*)
{endregion}
FUNCTION_BLOCK AssertArrayAllEqual_Byte EXTENDS AssertionBase
VAR_INPUT
    StartIndex : DINT; //! First selected index in IN; uses the array's declared index range, not a zero-based offset.
    Length : USINT; //! Number of compared elements, from 1 through 255.
    Expected : BYTE; //! Reference value for comparison with IN.
    Mask : BYTE := BYTE#16#FF; //! Bits included in the comparison; bits outside the mask are ignored.
END_VAR
VAR_IN_OUT CONSTANT
    IN : ARRAY[*] OF BYTE; //! Read-only compared data; keep stable during the call.
END_VAR

SUPER^();

{region 'Documentation'}
(*!
<summary>Validate configuration before comparing the selected range.</summary>
*)
{endregion}
METHOD PROTECTED Assert
VAR
    InLowerIndex : DINT;
    InUpperIndex : DINT;
    EndIndex : LINT;
    Offset : LINT;
    InIndex : DINT;
    ValuesEqual : BOOL;
    Message : STRING(GVL_Constants.MessageLength);
    ActualText : STRING(GVL_Constants.AssertionValueLength);
    ExpectedText : STRING(GVL_Constants.AssertionValueLength);
END_VAR
VAR CONSTANT
    HexDigitCount : USINT := 2;
END_VAR
IF NOT EvaluationActive THEN
    RETURN;
END_IF;

IF Result = E_Result.Error THEN
    RETURN;
END_IF;

// C0371: FB input is checked here before any reference access.
{warning disable C0371}
IF NOT __ISVALIDREF(IN) THEN
    Error(Message := 'Assertion error: IN reference is invalid.');
    RETURN;
END_IF;

InLowerIndex := LOWER_BOUND(IN, 1);
InUpperIndex := UPPER_BOUND(IN, 1);
EndIndex := DINT_TO_LINT(StartIndex) + USINT_TO_LINT(Length) - 1;

IF (Length = 0)
    OR (StartIndex < InLowerIndex) OR (StartIndex > InUpperIndex)
    OR (EndIndex > DINT_TO_LINT(InUpperIndex)) THEN
    Message := CONCAT('Assertion error: array range is invalid. StartIndex = ',
        DINT_TO_STRING(StartIndex));
    Message := CONCAT(Message, ', Length = ');
    Message := CONCAT(Message, USINT_TO_STRING(Length));
    Message := CONCAT(Message, '.');
    Error(Message := Message);
    RETURN;
END_IF;

IF Result = E_Result.Failed THEN
    RETURN;
END_IF;

FOR Offset := 0 TO USINT_TO_LINT(Length) - 1 DO
    InIndex := LINT_TO_DINT(DINT_TO_LINT(StartIndex) + Offset);
    ValuesEqual := FALSE;
    ValuesEqual := (IN[InIndex] AND Mask) = (Expected AND Mask);
    IF NOT ValuesEqual THEN
        EXIT;
    END_IF;
END_FOR;

IF NOT ValuesEqual THEN
    ExpectedText := CreateAssertionTextValue_Hex(Value := BYTE_TO_LWORD(Expected),
        DigitCount := HexDigitCount);
    ActualText := CreateAssertionTextValue_Hex(Value := BYTE_TO_LWORD(IN[InIndex]),
        DigitCount := HexDigitCount);
    Message := CONCAT('Assertion failed: array value is not equal. Expected = ',
        ExpectedText);
    Message := CONCAT(Message, ', Actual[');
    Message := CONCAT(Message, DINT_TO_STRING(InIndex));
    Message := CONCAT(Message, '] = ');
    Message := CONCAT(Message, ActualText);
    Message := CONCAT(Message, ', Range = [');
    Message := CONCAT(Message, DINT_TO_STRING(StartIndex));
    Message := CONCAT(Message, '..');
    Message := CONCAT(Message, LINT_TO_STRING(EndIndex));
    Message := CONCAT(Message, ']');
    Message := CONCAT(Message, ', Mask = ');
    Message := CONCAT(Message, CreateAssertionTextValue_Hex(Value := BYTE_TO_LWORD(Mask),
        DigitCount := HexDigitCount));
    Message := CONCAT(Message, '.');
    Fail(Message := Message);
    RETURN;
END_IF;

Pass();
{warning restore C0371}
END_METHOD

END_FUNCTION_BLOCK

// ---- Framework/Assertions/POU/Arrays/Byte/AssertArrayContainsArray_Byte.TcPOU
{region 'Documentation'}
(*!
<summary>Searches the selected IN range for the complete contiguous Expected pattern.</summary>
<description>

StartIndex is an absolute declared IN index, not an offset. Length selects 1..255
elements; the complete selected range must fit IN. Invalid references or ranges report
Error.

Keep supplied arrays stable for the call. Input data is read, not copied or retained as a
snapshot.

Comparison applies Mask to both values; bits outside it are ignored. The default mask
selects all bits.

The complete Expected pattern must be nonempty and fit the selected IN range; an
oversized pattern reports Error, not a missing-match result.

</description>
*)
{endregion}
FUNCTION_BLOCK AssertArrayContainsArray_Byte EXTENDS AssertionBase
VAR_INPUT
    StartIndex : DINT; //! First selected index in IN; uses the array's declared index range, not a zero-based offset.
    Length : USINT; //! Number of searched elements, from 1 through 255.
    Mask : BYTE := BYTE#16#FF; //! Bits included in the comparison; bits outside the mask are ignored.
END_VAR
VAR_IN_OUT CONSTANT
    IN : ARRAY[*] OF BYTE; //! Read-only search data; keep stable during the call.
    Expected : ARRAY[*] OF BYTE; //! Read-only expected sequence starting at its own lower bound; must fit the selected actual range.
END_VAR

SUPER^();

{region 'Documentation'}
(*!
<summary>Validate configuration before searching the selected range.</summary>
*)
{endregion}
METHOD PROTECTED Assert
VAR
    InLowerIndex : DINT;
    InUpperIndex : DINT;
    EndIndex : LINT;
    Offset : LINT;
    InIndex : DINT;
    ExpectedLowerIndex : DINT;
    ExpectedUpperIndex : DINT;
    ExpectedLength : LINT;
    ExpectedIndex : DINT;
    CandidateOffset : LINT;
    PatternFound : BOOL;
    PatternMatches : BOOL;
    Message : STRING(GVL_Constants.MessageLength);
END_VAR
VAR CONSTANT
    HexDigitCount : USINT := 2;
END_VAR
IF NOT EvaluationActive THEN
    RETURN;
END_IF;

IF Result = E_Result.Error THEN
    RETURN;
END_IF;

// C0371: FB input is checked here before any reference access.
{warning disable C0371}
IF NOT __ISVALIDREF(IN) THEN
    Error(Message := 'Assertion error: IN reference is invalid.');
    RETURN;
END_IF;

IF NOT __ISVALIDREF(Expected) THEN
    Error(Message := 'Assertion error: Expected reference is invalid.');
    RETURN;
END_IF;

InLowerIndex := LOWER_BOUND(IN, 1);
InUpperIndex := UPPER_BOUND(IN, 1);
EndIndex := DINT_TO_LINT(StartIndex) + USINT_TO_LINT(Length) - 1;

ExpectedLowerIndex := LOWER_BOUND(Expected, 1);
ExpectedUpperIndex := UPPER_BOUND(Expected, 1);
ExpectedLength := DINT_TO_LINT(ExpectedUpperIndex) - DINT_TO_LINT(ExpectedLowerIndex) + 1;

IF (Length = 0)
    OR (ExpectedLength <= 0) OR (ExpectedLength > USINT_TO_LINT(Length))
    OR (StartIndex < InLowerIndex) OR (StartIndex > InUpperIndex)
    OR (EndIndex > DINT_TO_LINT(InUpperIndex)) THEN
    Message := CONCAT('Assertion error: array range or pattern is invalid. StartIndex = ',
        DINT_TO_STRING(StartIndex));
    Message := CONCAT(Message, ', Length = ');
    Message := CONCAT(Message, USINT_TO_STRING(Length));
    Message := CONCAT(Message, ', ExpectedLength = ');
    Message := CONCAT(Message, LINT_TO_STRING(ExpectedLength));
    Message := CONCAT(Message, '.');
    Error(Message := Message);
    RETURN;
END_IF;

IF Result = E_Result.Failed THEN
    RETURN;
END_IF;

PatternFound := FALSE;
FOR CandidateOffset := 0 TO USINT_TO_LINT(Length) - ExpectedLength DO
    PatternMatches := TRUE;
    FOR Offset := 0 TO ExpectedLength - 1 DO
        InIndex := LINT_TO_DINT(DINT_TO_LINT(StartIndex) + CandidateOffset + Offset);
        ExpectedIndex := LINT_TO_DINT(DINT_TO_LINT(ExpectedLowerIndex) + Offset);
        IF (IN[InIndex] AND Mask) <> (Expected[ExpectedIndex] AND Mask) THEN
            PatternMatches := FALSE;
            EXIT;
        END_IF;
    END_FOR;

    IF PatternMatches THEN
        PatternFound := TRUE;
        EXIT;
    END_IF;
END_FOR;

IF NOT PatternFound THEN
    Message := CONCAT('Assertion failed: array range does not contain Expected pattern. ExpectedRange = [',
        DINT_TO_STRING(ExpectedLowerIndex));
    Message := CONCAT(Message, '..');
    Message := CONCAT(Message, DINT_TO_STRING(ExpectedUpperIndex));
    Message := CONCAT(Message, '], ActualRange = [');
    Message := CONCAT(Message, DINT_TO_STRING(StartIndex));
    Message := CONCAT(Message, '..');
    Message := CONCAT(Message, LINT_TO_STRING(EndIndex));
    Message := CONCAT(Message, ']');
    Message := CONCAT(Message, ', Mask = ');
    Message := CONCAT(Message, CreateAssertionTextValue_Hex(Value := BYTE_TO_LWORD(Mask),
        DigitCount := HexDigitCount));
    Message := CONCAT(Message, '.');
    Fail(Message := Message);
    RETURN;
END_IF;

Pass();
{warning restore C0371}
END_METHOD

END_FUNCTION_BLOCK

// ---- Framework/Assertions/POU/Arrays/Byte/AssertArrayContainsValue_Byte.TcPOU
{region 'Documentation'}
(*!
<summary>Searches the selected IN range for Expected; invalid configuration reports
Error.</summary>
<description>

StartIndex is an absolute declared IN index, not an offset. Length selects 1..255
elements; the complete selected range must fit IN. Invalid references or ranges report
Error.

Keep supplied arrays stable for the call. Input data is read, not copied or retained as a
snapshot.

Comparison applies Mask to both values; bits outside it are ignored. The default mask
selects all bits.

</description>
*)
{endregion}
FUNCTION_BLOCK AssertArrayContainsValue_Byte EXTENDS AssertionBase
VAR_INPUT
    StartIndex : DINT; //! First selected index in IN; uses the array's declared index range, not a zero-based offset.
    Length : USINT; //! Number of searched elements, from 1 through 255.
    Expected : BYTE; //! Reference value for comparison with IN.
    Mask : BYTE := BYTE#16#FF; //! Bits included in the comparison; bits outside the mask are ignored.
END_VAR
VAR_IN_OUT CONSTANT
    IN : ARRAY[*] OF BYTE; //! Read-only search data; keep stable during the call.
END_VAR

SUPER^();

{region 'Documentation'}
(*!
<summary>Validate configuration before searching the selected range.</summary>
*)
{endregion}
METHOD PROTECTED Assert
VAR
    InLowerIndex : DINT;
    InUpperIndex : DINT;
    EndIndex : LINT;
    Offset : LINT;
    InIndex : DINT;
    ValueFound : BOOL;
    Message : STRING(GVL_Constants.MessageLength);
    ExpectedText : STRING(GVL_Constants.AssertionValueLength);
END_VAR
VAR CONSTANT
    HexDigitCount : USINT := 2;
END_VAR
IF NOT EvaluationActive THEN
    RETURN;
END_IF;

IF Result = E_Result.Error THEN
    RETURN;
END_IF;

// C0371: FB input is checked here before any reference access.
{warning disable C0371}
IF NOT __ISVALIDREF(IN) THEN
    Error(Message := 'Assertion error: IN reference is invalid.');
    RETURN;
END_IF;

InLowerIndex := LOWER_BOUND(IN, 1);
InUpperIndex := UPPER_BOUND(IN, 1);
EndIndex := DINT_TO_LINT(StartIndex) + USINT_TO_LINT(Length) - 1;

IF (Length = 0)
    OR (StartIndex < InLowerIndex) OR (StartIndex > InUpperIndex)
    OR (EndIndex > DINT_TO_LINT(InUpperIndex)) THEN
    Message := CONCAT('Assertion error: array range is invalid. StartIndex = ',
        DINT_TO_STRING(StartIndex));
    Message := CONCAT(Message, ', Length = ');
    Message := CONCAT(Message, USINT_TO_STRING(Length));
    Message := CONCAT(Message, '.');
    Error(Message := Message);
    RETURN;
END_IF;

IF Result = E_Result.Failed THEN
    RETURN;
END_IF;

ValueFound := FALSE;
FOR Offset := 0 TO USINT_TO_LINT(Length) - 1 DO
    InIndex := LINT_TO_DINT(DINT_TO_LINT(StartIndex) + Offset);
    ValueFound := (IN[InIndex] AND Mask) = (Expected AND Mask);
    IF ValueFound THEN
        EXIT;
    END_IF;
END_FOR;

IF NOT ValueFound THEN
    ExpectedText := CreateAssertionTextValue_Hex(Value := BYTE_TO_LWORD(Expected),
        DigitCount := HexDigitCount);
    Message := CONCAT('Assertion failed: array range does not contain Expected = ',
        ExpectedText);
    Message := CONCAT(Message, ', Range = [');
    Message := CONCAT(Message, DINT_TO_STRING(StartIndex));
    Message := CONCAT(Message, '..');
    Message := CONCAT(Message, LINT_TO_STRING(EndIndex));
    Message := CONCAT(Message, ']');
    Message := CONCAT(Message, ', Mask = ');
    Message := CONCAT(Message, CreateAssertionTextValue_Hex(Value := BYTE_TO_LWORD(Mask),
        DigitCount := HexDigitCount));
    Message := CONCAT(Message, '.');
    Fail(Message := Message);
    RETURN;
END_IF;

Pass();
{warning restore C0371}
END_METHOD

END_FUNCTION_BLOCK

// ---- Framework/Assertions/POU/Arrays/Byte/AssertArrayEndsWithArray_Byte.TcPOU
{region 'Documentation'}
(*!
<summary>Compares Expected with the suffix of the selected IN range.</summary>
<description>

StartIndex is an absolute declared IN index, not an offset. Length selects 1..255
elements; the complete selected range must fit IN. Invalid references or ranges report
Error.

Keep supplied arrays stable for the call. Input data is read, not copied or retained as a
snapshot.

Comparison applies Mask to both values; bits outside it are ignored. The default mask
selects all bits.

The complete Expected pattern must be nonempty and fit the selected IN range; an
oversized pattern reports Error, not a missing-match result.

</description>
*)
{endregion}
FUNCTION_BLOCK AssertArrayEndsWithArray_Byte EXTENDS AssertionBase
VAR_INPUT
    Mask : BYTE := BYTE#16#FF; //! Bits included in each element comparison.
    StartIndex : DINT; //! First index of the selected IN range.
    Length : USINT; //! Number of selected elements starting at StartIndex; must fit the array range; valid range 1..255.
END_VAR
VAR_IN_OUT CONSTANT
    IN : ARRAY[*] OF BYTE; //! Read-only actual data; the selected range must remain stable during the call.
    Expected : ARRAY[*] OF BYTE; //! Read-only expected sequence starting at its own lower bound; must fit the selected actual range.
END_VAR

SUPER^();

{region 'Documentation'}
(*!
<summary>Validate the selected range and expectations before comparing elements.</summary>
*)
{endregion}
METHOD PROTECTED Assert
VAR
    InLowerIndex : DINT;
    InUpperIndex : DINT;
    ExpectedLowerIndex : DINT;
    ExpectedUpperIndex : DINT;
    ExpectedLength : LINT;
    EndIndex : LINT;
    Offset : LINT;
    InIndex : DINT;
    ExpectedIndex : DINT;
    Message : STRING(GVL_Constants.MessageLength);
    ExpectedText : STRING(GVL_Constants.AssertionValueLength);
    ActualText : STRING(GVL_Constants.AssertionValueLength);
END_VAR
VAR CONSTANT
    HexDigitCount : USINT := 2;
END_VAR
IF NOT EvaluationActive THEN
    RETURN;
END_IF;

IF Result = E_Result.Error THEN
    RETURN;
END_IF;

// C0371: FB inputs are checked here before any reference access.
{warning disable C0371}
IF NOT __ISVALIDREF(IN) THEN
    Error(Message := 'Assertion error: IN reference is invalid.');
    RETURN;
END_IF;

IF NOT __ISVALIDREF(Expected) THEN
    Error(Message := 'Assertion error: Expected reference is invalid.');
    RETURN;
END_IF;

InLowerIndex := LOWER_BOUND(IN, 1);
InUpperIndex := UPPER_BOUND(IN, 1);
ExpectedLowerIndex := LOWER_BOUND(Expected, 1);
ExpectedUpperIndex := UPPER_BOUND(Expected, 1);
ExpectedLength := DINT_TO_LINT(ExpectedUpperIndex) - DINT_TO_LINT(ExpectedLowerIndex) + 1;
EndIndex := DINT_TO_LINT(StartIndex) + USINT_TO_LINT(Length) - 1;

IF (Length = 0) OR (ExpectedLength <= 0)
    OR (ExpectedLength > USINT_TO_LINT(Length))
    OR (StartIndex < InLowerIndex) OR (StartIndex > InUpperIndex)
    OR (EndIndex > DINT_TO_LINT(InUpperIndex)) THEN
    Message := CONCAT('Assertion error: array range is invalid. StartIndex = ',
        DINT_TO_STRING(StartIndex));
    Message := CONCAT(Message, ', EndIndex = ');
    Message := CONCAT(Message, LINT_TO_STRING(EndIndex));
    Message := CONCAT(Message, ', InLowerIndex = ');
    Message := CONCAT(Message, DINT_TO_STRING(InLowerIndex));
    Message := CONCAT(Message, ', InUpperIndex = ');
    Message := CONCAT(Message, DINT_TO_STRING(InUpperIndex));
    Message := CONCAT(Message, ', ExpectedLength = ');
    Message := CONCAT(Message, LINT_TO_STRING(ExpectedLength));
    Message := CONCAT(Message, '.');
    Error(Message := Message);
    RETURN;
END_IF;

IF Result = E_Result.Failed THEN
    RETURN;
END_IF;

FOR Offset := 0 TO ExpectedLength - 1 DO
    InIndex := LINT_TO_DINT(EndIndex - ExpectedLength + 1 + Offset);
    ExpectedIndex := LINT_TO_DINT(DINT_TO_LINT(ExpectedLowerIndex) + Offset);
    IF (IN[InIndex] AND Mask) <> (Expected[ExpectedIndex] AND Mask) THEN
        ExpectedText := CreateAssertionTextValue_Hex(Value := BYTE_TO_LWORD(Expected[ExpectedIndex]),
            DigitCount := HexDigitCount);
        ActualText := CreateAssertionTextValue_Hex(Value := BYTE_TO_LWORD(IN[InIndex]),
            DigitCount := HexDigitCount);
        Message := CONCAT('Assertion failed: array suffix differs. Expected[',
            DINT_TO_STRING(ExpectedIndex));
        Message := CONCAT(Message, '] = ');
        Message := CONCAT(Message, ExpectedText);
        Message := CONCAT(Message, ', IN[');
        Message := CONCAT(Message, DINT_TO_STRING(InIndex));
        Message := CONCAT(Message, '] = ');
        Message := CONCAT(Message, ActualText);
        Message := CONCAT(Message, '.');
        Message := CONCAT(Message, ' Mask = ');
        Message := CONCAT(Message, CreateAssertionTextValue_Hex(Value := BYTE_TO_LWORD(Mask),
            DigitCount := HexDigitCount));
        Fail(Message := Message);
        RETURN;
    END_IF;
END_FOR;

Pass();
{warning restore C0371}
END_METHOD

END_FUNCTION_BLOCK

// ---- Framework/Assertions/POU/Arrays/Byte/AssertArrayNoValueChange_Byte.TcPOU
{region 'Documentation'}
(*!
<summary>Captures one snapshot until Reset; Disable/Re-Enable never replaces it.</summary>
<description>

Disabling observation preserves the original snapshot. Re-enabling requires a fresh
preceding observation before comparisons resume; it does not replace that snapshot.

StartIndex is an absolute IN index and Length selects 1..255 elements within IN. Memory
must have at least Length elements from its own lower bound. Invalid references or ranges
report Error.

The caller provides dedicated writable Memory that must not overlap IN; overlap is not
checked. Keep bindings, selected range and snapshot contents stable until Reset. Reset
invalidates the snapshot without clearing Memory bytes.

</description>
*)
{endregion}
FUNCTION_BLOCK AssertArrayNoValueChange_Byte EXTENDS AssertionBase
VAR_INPUT
    Mask : BYTE := BYTE#16#FF; //! Bits included in each element comparison.
    StartIndex : DINT; //! First selected index in IN; uses the array's declared index range, not a zero-based offset.
    Length : USINT; //! Number of monitored elements, from 1 through 255.
END_VAR
VAR_IN_OUT CONSTANT
    IN : ARRAY[*] OF BYTE; //! Read-only actual data; the selected range must remain stable during the call.
END_VAR
VAR_IN_OUT
    Memory : ARRAY[*] OF BYTE; //! Dedicated snapshot storage; only this assertion writes its selected elements.
END_VAR
VAR
    FSnapshotValid : BOOL;
    FObservationPrevious : BOOL;
    FEvaluationActive : BOOL;
END_VAR

SUPER^();

{region 'Documentation'}
(*!
<summary>Capture once or compare against the retained snapshot after range validation.</summary>
*)
{endregion}
METHOD PROTECTED Assert
VAR
    InLowerIndex : DINT;
    InUpperIndex : DINT;
    MemoryLowerIndex : DINT;
    MemoryUpperIndex : DINT;
    MemoryEndIndex : LINT;
    EndIndex : LINT;
    Offset : LINT;
    InIndex : DINT;
    MemoryIndex : DINT;
    Message : STRING(GVL_Constants.MessageLength);
    ReferenceText : STRING(GVL_Constants.AssertionValueLength);
    ActualText : STRING(GVL_Constants.AssertionValueLength);
END_VAR
VAR CONSTANT
    HexDigitCount : USINT := 2;
END_VAR
FEvaluationActive := ObservationActive AND FObservationPrevious AND FSnapshotValid;
FObservationPrevious := ObservationActive;

IF NOT ObservationActive THEN
    RETURN;
END_IF;

IF Result = E_Result.Error THEN
    RETURN;
END_IF;

// C0371: FB inputs are checked here before any reference access.
{warning disable C0371}
IF NOT __ISVALIDREF(IN) THEN
    Error(Message := 'Assertion error: IN reference is invalid.');
    RETURN;
END_IF;

IF NOT __ISVALIDREF(Memory) THEN
    Error(Message := 'Assertion error: Memory reference is invalid.');
    RETURN;
END_IF;

InLowerIndex := LOWER_BOUND(IN, 1);
InUpperIndex := UPPER_BOUND(IN, 1);
MemoryLowerIndex := LOWER_BOUND(Memory, 1);
MemoryUpperIndex := UPPER_BOUND(Memory, 1);
EndIndex := DINT_TO_LINT(StartIndex) + USINT_TO_LINT(Length) - 1;
MemoryEndIndex := DINT_TO_LINT(MemoryLowerIndex) + USINT_TO_LINT(Length) - 1;

IF (Length = 0)
    OR (StartIndex < InLowerIndex) OR (StartIndex > InUpperIndex)
    OR (EndIndex > DINT_TO_LINT(InUpperIndex))
    OR (MemoryEndIndex > DINT_TO_LINT(MemoryUpperIndex)) THEN
    Message := CONCAT('Assertion error: array or memory range is invalid. StartIndex = ',
        DINT_TO_STRING(StartIndex));
    Message := CONCAT(Message, ', EndIndex = ');
    Message := CONCAT(Message, LINT_TO_STRING(EndIndex));
    Message := CONCAT(Message, ', Length = ');
    Message := CONCAT(Message, USINT_TO_STRING(Length));
    Message := CONCAT(Message, '.');
    Error(Message := Message);
    RETURN;
END_IF;

IF NOT FSnapshotValid THEN
    FOR Offset := 0 TO USINT_TO_LINT(Length) - 1 DO
        InIndex := LINT_TO_DINT(DINT_TO_LINT(StartIndex) + Offset);
        MemoryIndex := LINT_TO_DINT(DINT_TO_LINT(MemoryLowerIndex) + Offset);
        Memory[MemoryIndex] := IN[InIndex];
    END_FOR;
    FSnapshotValid := TRUE;
    RETURN;
END_IF;

IF NOT EvaluationActive THEN
    RETURN;
END_IF;

IF Result = E_Result.Failed THEN
    RETURN;
END_IF;

FOR Offset := 0 TO USINT_TO_LINT(Length) - 1 DO
    InIndex := LINT_TO_DINT(DINT_TO_LINT(StartIndex) + Offset);
    MemoryIndex := LINT_TO_DINT(DINT_TO_LINT(MemoryLowerIndex) + Offset);
    IF (IN[InIndex] AND Mask) <> (Memory[MemoryIndex] AND Mask) THEN
        ReferenceText := CreateAssertionTextValue_Hex(Value := BYTE_TO_LWORD(Memory[MemoryIndex]),
            DigitCount := HexDigitCount);
        ActualText := CreateAssertionTextValue_Hex(Value := BYTE_TO_LWORD(IN[InIndex]),
            DigitCount := HexDigitCount);
        Message := CONCAT('Assertion failed: array value changed. Reference[',
            DINT_TO_STRING(MemoryIndex));
        Message := CONCAT(Message, '] = ');
        Message := CONCAT(Message, ReferenceText);
        Message := CONCAT(Message, ', IN[');
        Message := CONCAT(Message, DINT_TO_STRING(InIndex));
        Message := CONCAT(Message, '] = ');
        Message := CONCAT(Message, ActualText);
        Message := CONCAT(Message, '.');
        Message := CONCAT(Message, ' Mask = ');
        Message := CONCAT(Message, CreateAssertionTextValue_Hex(Value := BYTE_TO_LWORD(Mask),
            DigitCount := HexDigitCount));
        Fail(Message := Message);
        RETURN;
    END_IF;
END_FOR;

Pass();
{warning restore C0371}
END_METHOD

{region 'Documentation'}
(*!
<summary>Current/last call has consecutive observation and an existing snapshot.</summary>
*)
{endregion}
{attribute 'monitoring' := 'call'}
PROPERTY PUBLIC EvaluationActive : BOOL //! Current/last call has consecutive observation and an existing snapshot.
GET // PUBLIC
EvaluationActive := FEvaluationActive;
END_GET
END_PROPERTY

{region 'Documentation'}
(*!
<summary>Invalidate the snapshot and observation history.</summary>
<description>

Does not clear external Memory. The next active observation captures a new snapshot
before comparison.

</description>
*)
{endregion}
METHOD PROTECTED ResetAssertion
FSnapshotValid := FALSE;
FObservationPrevious := FALSE;
FEvaluationActive := FALSE;
END_METHOD

END_FUNCTION_BLOCK

// ---- Framework/Assertions/POU/Arrays/Char/AssertArrayAllEqual_Char.TcPOU
{region 'Documentation'}
(*!
<summary>Character codes use BYTE; exact comparison without a mask.</summary>
<description>

Checks every selected IN element against Expected; reports the first mismatch.

StartIndex is an absolute declared IN index, not an offset. Length selects 1..255
elements; the complete selected range must fit IN. Invalid references or ranges report
Error.

Keep supplied arrays stable for the call. Input data is read, not copied or retained as a
snapshot.

</description>
*)
{endregion}
FUNCTION_BLOCK AssertArrayAllEqual_Char EXTENDS AssertionBase
VAR_INPUT
    StartIndex : DINT; //! First selected index in IN; uses the array's declared index range, not a zero-based offset.
    Length : USINT; //! Number of compared elements, from 1 through 255.
    Expected : BYTE; //! Reference value for comparison with IN.
END_VAR
VAR_IN_OUT CONSTANT
    IN : ARRAY[*] OF BYTE; //! Read-only compared data; keep stable during the call.
END_VAR

SUPER^();

{region 'Documentation'}
(*!
<summary>Validate configuration before comparing the selected range.</summary>
*)
{endregion}
METHOD PROTECTED Assert
VAR
    InLowerIndex : DINT;
    InUpperIndex : DINT;
    EndIndex : LINT;
    Offset : LINT;
    InIndex : DINT;
    ValuesEqual : BOOL;
    Message : STRING(GVL_Constants.MessageLength);
    ActualText : STRING;
    ExpectedText : STRING;
END_VAR
IF NOT EvaluationActive THEN
    RETURN;
END_IF;

IF Result = E_Result.Error THEN
    RETURN;
END_IF;

// C0371: FB input is checked here before any reference access.
{warning disable C0371}
IF NOT __ISVALIDREF(IN) THEN
    Error(Message := 'Assertion error: IN reference is invalid.');
    RETURN;
END_IF;

InLowerIndex := LOWER_BOUND(IN, 1);
InUpperIndex := UPPER_BOUND(IN, 1);
EndIndex := DINT_TO_LINT(StartIndex) + USINT_TO_LINT(Length) - 1;

IF (Length = 0)
    OR (StartIndex < InLowerIndex) OR (StartIndex > InUpperIndex)
    OR (EndIndex > DINT_TO_LINT(InUpperIndex)) THEN
    Message := CONCAT('Assertion error: array range is invalid. StartIndex = ',
        DINT_TO_STRING(StartIndex));
    Message := CONCAT(Message, ', Length = ');
    Message := CONCAT(Message, USINT_TO_STRING(Length));
    Message := CONCAT(Message, '.');
    Error(Message := Message);
    RETURN;
END_IF;

IF Result = E_Result.Failed THEN
    RETURN;
END_IF;

FOR Offset := 0 TO USINT_TO_LINT(Length) - 1 DO
    InIndex := LINT_TO_DINT(DINT_TO_LINT(StartIndex) + Offset);
    ValuesEqual := FALSE;
    ValuesEqual := IN[InIndex] = Expected;
    IF NOT ValuesEqual THEN
        EXIT;
    END_IF;
END_FOR;

IF NOT ValuesEqual THEN
    ExpectedText := CreateAssertionTextValue_Char(Value := Expected);
    ActualText := CreateAssertionTextValue_Char(Value := IN[InIndex]);
    Message := CONCAT('Assertion failed: array value is not equal. Expected = ',
        ExpectedText);
    Message := CONCAT(Message, ', Actual[');
    Message := CONCAT(Message, DINT_TO_STRING(InIndex));
    Message := CONCAT(Message, '] = ');
    Message := CONCAT(Message, ActualText);
    Message := CONCAT(Message, ', Range = [');
    Message := CONCAT(Message, DINT_TO_STRING(StartIndex));
    Message := CONCAT(Message, '..');
    Message := CONCAT(Message, LINT_TO_STRING(EndIndex));
    Message := CONCAT(Message, ']');
    Message := CONCAT(Message, '.');
    Fail(Message := Message);
    RETURN;
END_IF;

Pass();
{warning restore C0371}
END_METHOD

END_FUNCTION_BLOCK

// ---- Framework/Assertions/POU/Arrays/Char/AssertArrayContainsArray_Char.TcPOU
{region 'Documentation'}
(*!
<summary>Character codes use BYTE; exact comparison without a mask.</summary>
<description>

Searches the selected IN range for the complete contiguous Expected pattern.

StartIndex is an absolute declared IN index, not an offset. Length selects 1..255
elements; the complete selected range must fit IN. Invalid references or ranges report
Error.

Keep supplied arrays stable for the call. Input data is read, not copied or retained as a
snapshot.

The complete Expected pattern must be nonempty and fit the selected IN range; an
oversized pattern reports Error, not a missing-match result.

</description>
*)
{endregion}
FUNCTION_BLOCK AssertArrayContainsArray_Char EXTENDS AssertionBase
VAR_INPUT
    StartIndex : DINT; //! First selected index in IN; uses the array's declared index range, not a zero-based offset.
    Length : USINT; //! Number of searched elements, from 1 through 255.
END_VAR
VAR_IN_OUT CONSTANT
    IN : ARRAY[*] OF BYTE; //! Read-only search data; keep stable during the call.
    Expected : ARRAY[*] OF BYTE; //! Read-only expected sequence starting at its own lower bound; must fit the selected actual range.
END_VAR

SUPER^();

{region 'Documentation'}
(*!
<summary>Validate configuration before searching the selected range.</summary>
*)
{endregion}
METHOD PROTECTED Assert
VAR
    InLowerIndex : DINT;
    InUpperIndex : DINT;
    EndIndex : LINT;
    Offset : LINT;
    InIndex : DINT;
    ExpectedLowerIndex : DINT;
    ExpectedUpperIndex : DINT;
    ExpectedLength : LINT;
    ExpectedIndex : DINT;
    CandidateOffset : LINT;
    PatternFound : BOOL;
    PatternMatches : BOOL;
    Message : STRING(GVL_Constants.MessageLength);
END_VAR
IF NOT EvaluationActive THEN
    RETURN;
END_IF;

IF Result = E_Result.Error THEN
    RETURN;
END_IF;

// C0371: FB input is checked here before any reference access.
{warning disable C0371}
IF NOT __ISVALIDREF(IN) THEN
    Error(Message := 'Assertion error: IN reference is invalid.');
    RETURN;
END_IF;

IF NOT __ISVALIDREF(Expected) THEN
    Error(Message := 'Assertion error: Expected reference is invalid.');
    RETURN;
END_IF;

InLowerIndex := LOWER_BOUND(IN, 1);
InUpperIndex := UPPER_BOUND(IN, 1);
EndIndex := DINT_TO_LINT(StartIndex) + USINT_TO_LINT(Length) - 1;

ExpectedLowerIndex := LOWER_BOUND(Expected, 1);
ExpectedUpperIndex := UPPER_BOUND(Expected, 1);
ExpectedLength := DINT_TO_LINT(ExpectedUpperIndex) - DINT_TO_LINT(ExpectedLowerIndex) + 1;

IF (Length = 0)
    OR (ExpectedLength <= 0) OR (ExpectedLength > USINT_TO_LINT(Length))
    OR (StartIndex < InLowerIndex) OR (StartIndex > InUpperIndex)
    OR (EndIndex > DINT_TO_LINT(InUpperIndex)) THEN
    Message := CONCAT('Assertion error: array range or pattern is invalid. StartIndex = ',
        DINT_TO_STRING(StartIndex));
    Message := CONCAT(Message, ', Length = ');
    Message := CONCAT(Message, USINT_TO_STRING(Length));
    Message := CONCAT(Message, ', ExpectedLength = ');
    Message := CONCAT(Message, LINT_TO_STRING(ExpectedLength));
    Message := CONCAT(Message, '.');
    Error(Message := Message);
    RETURN;
END_IF;

IF Result = E_Result.Failed THEN
    RETURN;
END_IF;

PatternFound := FALSE;
FOR CandidateOffset := 0 TO USINT_TO_LINT(Length) - ExpectedLength DO
    PatternMatches := TRUE;
    FOR Offset := 0 TO ExpectedLength - 1 DO
        InIndex := LINT_TO_DINT(DINT_TO_LINT(StartIndex) + CandidateOffset + Offset);
        ExpectedIndex := LINT_TO_DINT(DINT_TO_LINT(ExpectedLowerIndex) + Offset);
        IF IN[InIndex] <> Expected[ExpectedIndex] THEN
            PatternMatches := FALSE;
            EXIT;
        END_IF;
    END_FOR;

    IF PatternMatches THEN
        PatternFound := TRUE;
        EXIT;
    END_IF;
END_FOR;

IF NOT PatternFound THEN
    Message := CONCAT('Assertion failed: array range does not contain Expected pattern. ExpectedRange = [',
        DINT_TO_STRING(ExpectedLowerIndex));
    Message := CONCAT(Message, '..');
    Message := CONCAT(Message, DINT_TO_STRING(ExpectedUpperIndex));
    Message := CONCAT(Message, '], ActualRange = [');
    Message := CONCAT(Message, DINT_TO_STRING(StartIndex));
    Message := CONCAT(Message, '..');
    Message := CONCAT(Message, LINT_TO_STRING(EndIndex));
    Message := CONCAT(Message, ']');
    Message := CONCAT(Message, '.');
    Fail(Message := Message);
    RETURN;
END_IF;

Pass();
{warning restore C0371}
END_METHOD

END_FUNCTION_BLOCK

// ---- Framework/Assertions/POU/Arrays/Char/AssertArrayContainsString_Char.TcPOU
{region 'Documentation'}
(*!
<summary>Search the selected array for the contiguous STRING code units.</summary>
<description>

StartIndex is an absolute declared IN index, not an offset. Length selects 1..255
elements; the complete selected range must fit IN. Invalid references or ranges report
Error.

Keep supplied arrays stable for the call. Input data is read, not copied or retained as a
snapshot.

Expected must be nonempty and fit its configured text capacity (otherwise Error). A valid
text longer than the selected array region reports Failed. The array is not zero-terminated or
trimmed; matching is exact and case-sensitive.

</description>
*)
{endregion}
FUNCTION_BLOCK AssertArrayContainsString_Char EXTENDS AssertionBase
VAR_INPUT
    StartIndex : DINT; //! First selected index in IN; uses the array's declared index range, not a zero-based offset.
    Length : USINT; //! Number of selected array elements, from 1 through 255.
END_VAR
VAR_IN_OUT CONSTANT
    IN : ARRAY[*] OF BYTE; //! Read-only actual data; the selected range must remain stable during the call.
    Expected : STRING(Param_Assertions.AssertionStringLength); //! Nonempty expected text, terminated within the configured capacity; keep stable during the call.
END_VAR

SUPER^();

{region 'Documentation'}
(*!
<summary>Validate references and ranges before exact code-unit comparison.</summary>
*)
{endregion}
METHOD PROTECTED Assert
VAR
    InLowerIndex : DINT;
    InUpperIndex : DINT;
    EndIndex : LINT;
    ExpectedLength : DINT;
    CharacterIndex : DINT;
    InIndex : DINT;
    CandidateOffset : LINT;
    LastCandidateOffset : LINT;
    PatternMatches : BOOL;
    PatternFound : BOOL;
    ExpectedText : STRING(GVL_Constants.AssertionValueLength);
    Message : STRING(GVL_Constants.MessageLength);
END_VAR
VAR CONSTANT
    Terminator : BYTE := 0;
END_VAR
IF NOT EvaluationActive THEN
    RETURN;
END_IF;

IF Result = E_Result.Error THEN
    RETURN;
END_IF;

// C0371: FB inputs are checked before any reference access.
{warning disable C0371}
IF NOT __ISVALIDREF(IN) THEN
    Error(Message := 'Assertion error: IN reference is invalid.');
    RETURN;
END_IF;

IF NOT __ISVALIDREF(Expected) THEN
    Error(Message := 'Assertion error: Expected reference is invalid.');
    RETURN;
END_IF;

IF NOT IsAssertionStringLengthValid(Value := Expected) THEN
    Error(Message := 'Assertion error: Expected exceeds configured STRING length.');
    RETURN;
END_IF;

IF Expected[0] = Terminator THEN
    Error(Message := 'Assertion error: Expected must not be empty.');
    RETURN;
END_IF;

ExpectedLength := 0;
FOR CharacterIndex := 0 TO UINT_TO_DINT(Param_Assertions.AssertionStringLength) DO
    IF Expected[CharacterIndex] = Terminator THEN
        ExpectedLength := CharacterIndex;
        EXIT;
    END_IF;
END_FOR;

InLowerIndex := LOWER_BOUND(IN, 1);
InUpperIndex := UPPER_BOUND(IN, 1);
EndIndex := DINT_TO_LINT(StartIndex) + USINT_TO_LINT(Length) - 1;
IF (Length = 0)
    OR (StartIndex < InLowerIndex) OR (StartIndex > InUpperIndex)
    OR (EndIndex > DINT_TO_LINT(InUpperIndex)) THEN
    Message := CONCAT('Assertion error: array range is invalid. StartIndex = ',
        DINT_TO_STRING(StartIndex));
    Message := CONCAT(Message, ', Length = ');
    Message := CONCAT(Message, USINT_TO_STRING(Length));
    Error(Message := Message);
    RETURN;
END_IF;

IF Result = E_Result.Failed THEN
    RETURN;
END_IF;

PatternFound := FALSE;
IF ExpectedLength <= USINT_TO_DINT(Length) THEN
    LastCandidateOffset := USINT_TO_LINT(Length) - DINT_TO_LINT(ExpectedLength);
    FOR CandidateOffset := 0 TO LastCandidateOffset DO
        PatternMatches := TRUE;
        FOR CharacterIndex := 0 TO ExpectedLength - 1 DO
            InIndex := LINT_TO_DINT(DINT_TO_LINT(StartIndex) + CandidateOffset
                + DINT_TO_LINT(CharacterIndex));
            IF IN[InIndex] <> Expected[CharacterIndex] THEN
                PatternMatches := FALSE;
                EXIT;
            END_IF;
        END_FOR;
        IF PatternMatches THEN
            PatternFound := TRUE;
            EXIT;
        END_IF;
    END_FOR;
END_IF;

IF NOT PatternFound THEN
    ExpectedText := CreateAssertionTextValue_String(Value := Expected);
    Message := CONCAT('Assertion failed: selected array does not contain Expected = ',
        ExpectedText);
    Message := CONCAT(Message, ', Range = [');
    Message := CONCAT(Message, DINT_TO_STRING(StartIndex));
    Message := CONCAT(Message, '..');
    Message := CONCAT(Message, LINT_TO_STRING(EndIndex));
    Message := CONCAT(Message, '], ExpectedLength = ');
    Message := CONCAT(Message, DINT_TO_STRING(ExpectedLength));
    Message := CONCAT(Message, '.');
    Fail(Message := Message);
    RETURN;
END_IF;

Pass();
{warning restore C0371}
END_METHOD

END_FUNCTION_BLOCK

// ---- Framework/Assertions/POU/Arrays/Char/AssertArrayContainsValue_Char.TcPOU
{region 'Documentation'}
(*!
<summary>Character codes use BYTE; exact comparison without a mask.</summary>
<description>

Searches the selected IN range for Expected; invalid configuration reports Error.

StartIndex is an absolute declared IN index, not an offset. Length selects 1..255
elements; the complete selected range must fit IN. Invalid references or ranges report
Error.

Keep supplied arrays stable for the call. Input data is read, not copied or retained as a
snapshot.

</description>
*)
{endregion}
FUNCTION_BLOCK AssertArrayContainsValue_Char EXTENDS AssertionBase
VAR_INPUT
    StartIndex : DINT; //! First selected index in IN; uses the array's declared index range, not a zero-based offset.
    Length : USINT; //! Number of searched elements, from 1 through 255.
    Expected : BYTE; //! Reference value for comparison with IN.
END_VAR
VAR_IN_OUT CONSTANT
    IN : ARRAY[*] OF BYTE; //! Read-only search data; keep stable during the call.
END_VAR

SUPER^();

{region 'Documentation'}
(*!
<summary>Validate configuration before searching the selected range.</summary>
*)
{endregion}
METHOD PROTECTED Assert
VAR
    InLowerIndex : DINT;
    InUpperIndex : DINT;
    EndIndex : LINT;
    Offset : LINT;
    InIndex : DINT;
    ValueFound : BOOL;
    Message : STRING(GVL_Constants.MessageLength);
    ExpectedText : STRING;
END_VAR
IF NOT EvaluationActive THEN
    RETURN;
END_IF;

IF Result = E_Result.Error THEN
    RETURN;
END_IF;

// C0371: FB input is checked here before any reference access.
{warning disable C0371}
IF NOT __ISVALIDREF(IN) THEN
    Error(Message := 'Assertion error: IN reference is invalid.');
    RETURN;
END_IF;

InLowerIndex := LOWER_BOUND(IN, 1);
InUpperIndex := UPPER_BOUND(IN, 1);
EndIndex := DINT_TO_LINT(StartIndex) + USINT_TO_LINT(Length) - 1;

IF (Length = 0)
    OR (StartIndex < InLowerIndex) OR (StartIndex > InUpperIndex)
    OR (EndIndex > DINT_TO_LINT(InUpperIndex)) THEN
    Message := CONCAT('Assertion error: array range is invalid. StartIndex = ',
        DINT_TO_STRING(StartIndex));
    Message := CONCAT(Message, ', Length = ');
    Message := CONCAT(Message, USINT_TO_STRING(Length));
    Message := CONCAT(Message, '.');
    Error(Message := Message);
    RETURN;
END_IF;

IF Result = E_Result.Failed THEN
    RETURN;
END_IF;

ValueFound := FALSE;
FOR Offset := 0 TO USINT_TO_LINT(Length) - 1 DO
    InIndex := LINT_TO_DINT(DINT_TO_LINT(StartIndex) + Offset);
    ValueFound := IN[InIndex] = Expected;
    IF ValueFound THEN
        EXIT;
    END_IF;
END_FOR;

IF NOT ValueFound THEN
    ExpectedText := CreateAssertionTextValue_Char(Value := Expected);
    Message := CONCAT('Assertion failed: array range does not contain Expected = ',
        ExpectedText);
    Message := CONCAT(Message, ', Range = [');
    Message := CONCAT(Message, DINT_TO_STRING(StartIndex));
    Message := CONCAT(Message, '..');
    Message := CONCAT(Message, LINT_TO_STRING(EndIndex));
    Message := CONCAT(Message, ']');
    Message := CONCAT(Message, '.');
    Fail(Message := Message);
    RETURN;
END_IF;

Pass();
{warning restore C0371}
END_METHOD

END_FUNCTION_BLOCK

// ---- Framework/Assertions/POU/Arrays/Char/AssertArrayEndsWithString_Char.TcPOU
{region 'Documentation'}
(*!
<summary>Check that the selected array ends with the STRING code units.</summary>
<description>

StartIndex is an absolute declared IN index, not an offset. Length selects 1..255
elements; the complete selected range must fit IN. Invalid references or ranges report
Error.

Keep supplied arrays stable for the call. Input data is read, not copied or retained as a
snapshot.

Expected must be nonempty and fit its configured text capacity (otherwise Error). A valid
text longer than the selected array region reports Failed. The array is not zero-terminated or
trimmed; matching is exact and case-sensitive.

</description>
*)
{endregion}
FUNCTION_BLOCK AssertArrayEndsWithString_Char EXTENDS AssertionBase
VAR_INPUT
    StartIndex : DINT; //! First selected index in IN; uses the array's declared index range, not a zero-based offset.
    Length : USINT; //! Number of selected array elements, from 1 through 255.
END_VAR
VAR_IN_OUT CONSTANT
    IN : ARRAY[*] OF BYTE; //! Read-only actual data; the selected range must remain stable during the call.
    Expected : STRING(Param_Assertions.AssertionStringLength); //! Nonempty expected text, terminated within the configured capacity; keep stable during the call.
END_VAR

SUPER^();

{region 'Documentation'}
(*!
<summary>Validate references and ranges before exact code-unit comparison.</summary>
*)
{endregion}
METHOD PROTECTED Assert
VAR
    InLowerIndex : DINT;
    InUpperIndex : DINT;
    EndIndex : LINT;
    ExpectedLength : DINT;
    CharacterIndex : DINT;
    InIndex : DINT;
    CandidateOffset : LINT;
    LastCandidateOffset : LINT;
    PatternMatches : BOOL;
    PatternFound : BOOL;
    ExpectedText : STRING(GVL_Constants.AssertionValueLength);
    Message : STRING(GVL_Constants.MessageLength);
END_VAR
VAR CONSTANT
    Terminator : BYTE := 0;
END_VAR
IF NOT EvaluationActive THEN
    RETURN;
END_IF;

IF Result = E_Result.Error THEN
    RETURN;
END_IF;

// C0371: FB inputs are checked before any reference access.
{warning disable C0371}
IF NOT __ISVALIDREF(IN) THEN
    Error(Message := 'Assertion error: IN reference is invalid.');
    RETURN;
END_IF;

IF NOT __ISVALIDREF(Expected) THEN
    Error(Message := 'Assertion error: Expected reference is invalid.');
    RETURN;
END_IF;

IF NOT IsAssertionStringLengthValid(Value := Expected) THEN
    Error(Message := 'Assertion error: Expected exceeds configured STRING length.');
    RETURN;
END_IF;

IF Expected[0] = Terminator THEN
    Error(Message := 'Assertion error: Expected must not be empty.');
    RETURN;
END_IF;

ExpectedLength := 0;
FOR CharacterIndex := 0 TO UINT_TO_DINT(Param_Assertions.AssertionStringLength) DO
    IF Expected[CharacterIndex] = Terminator THEN
        ExpectedLength := CharacterIndex;
        EXIT;
    END_IF;
END_FOR;

InLowerIndex := LOWER_BOUND(IN, 1);
InUpperIndex := UPPER_BOUND(IN, 1);
EndIndex := DINT_TO_LINT(StartIndex) + USINT_TO_LINT(Length) - 1;
IF (Length = 0)
    OR (StartIndex < InLowerIndex) OR (StartIndex > InUpperIndex)
    OR (EndIndex > DINT_TO_LINT(InUpperIndex)) THEN
    Message := CONCAT('Assertion error: array range is invalid. StartIndex = ',
        DINT_TO_STRING(StartIndex));
    Message := CONCAT(Message, ', Length = ');
    Message := CONCAT(Message, USINT_TO_STRING(Length));
    Error(Message := Message);
    RETURN;
END_IF;

IF Result = E_Result.Failed THEN
    RETURN;
END_IF;

PatternFound := FALSE;
IF ExpectedLength <= USINT_TO_DINT(Length) THEN
    LastCandidateOffset := USINT_TO_LINT(Length) - DINT_TO_LINT(ExpectedLength);
    FOR CandidateOffset := USINT_TO_LINT(Length) - DINT_TO_LINT(ExpectedLength) TO LastCandidateOffset DO
        PatternMatches := TRUE;
        FOR CharacterIndex := 0 TO ExpectedLength - 1 DO
            InIndex := LINT_TO_DINT(DINT_TO_LINT(StartIndex) + CandidateOffset
                + DINT_TO_LINT(CharacterIndex));
            IF IN[InIndex] <> Expected[CharacterIndex] THEN
                PatternMatches := FALSE;
                EXIT;
            END_IF;
        END_FOR;
        IF PatternMatches THEN
            PatternFound := TRUE;
            EXIT;
        END_IF;
    END_FOR;
END_IF;

IF NOT PatternFound THEN
    ExpectedText := CreateAssertionTextValue_String(Value := Expected);
    Message := CONCAT('Assertion failed: selected array does not end with Expected = ',
        ExpectedText);
    Message := CONCAT(Message, ', Range = [');
    Message := CONCAT(Message, DINT_TO_STRING(StartIndex));
    Message := CONCAT(Message, '..');
    Message := CONCAT(Message, LINT_TO_STRING(EndIndex));
    Message := CONCAT(Message, '], ExpectedLength = ');
    Message := CONCAT(Message, DINT_TO_STRING(ExpectedLength));
    Message := CONCAT(Message, '.');
    Fail(Message := Message);
    RETURN;
END_IF;

Pass();
{warning restore C0371}
END_METHOD

END_FUNCTION_BLOCK

// ---- Framework/Assertions/POU/Arrays/Char/AssertArrayEqualString_Char.TcPOU
{region 'Documentation'}
(*!
<summary>Check that the selected array exactly equals the STRING code units.</summary>
<description>

StartIndex is an absolute declared IN index, not an offset. Length selects 1..255
elements; the complete selected range must fit IN. Invalid references or ranges report
Error.

Keep supplied arrays stable for the call. Input data is read, not copied or retained as a
snapshot.

Expected must be nonempty and fit its configured text capacity (otherwise Error). A valid
text longer than the selected array region reports Failed. The array is not zero-terminated or
trimmed; matching is exact and case-sensitive.

The selected array length must equal the text length; trailing padding counts as
data.

</description>
*)
{endregion}
FUNCTION_BLOCK AssertArrayEqualString_Char EXTENDS AssertionBase
VAR_INPUT
    StartIndex : DINT; //! First selected index in IN; uses the array's declared index range, not a zero-based offset.
    Length : USINT; //! Number of selected array elements, from 1 through 255.
END_VAR
VAR_IN_OUT CONSTANT
    IN : ARRAY[*] OF BYTE; //! Read-only actual data; the selected range must remain stable during the call.
    Expected : STRING(Param_Assertions.AssertionStringLength); //! Nonempty expected text, terminated within the configured capacity; keep stable during the call.
END_VAR

SUPER^();

{region 'Documentation'}
(*!
<summary>Validate references and ranges before exact code-unit comparison.</summary>
*)
{endregion}
METHOD PROTECTED Assert
VAR
    InLowerIndex : DINT;
    InUpperIndex : DINT;
    EndIndex : LINT;
    ExpectedLength : DINT;
    CharacterIndex : DINT;
    InIndex : DINT;
    CandidateOffset : LINT;
    LastCandidateOffset : LINT;
    PatternMatches : BOOL;
    PatternFound : BOOL;
    ExpectedText : STRING(GVL_Constants.AssertionValueLength);
    Message : STRING(GVL_Constants.MessageLength);
END_VAR
VAR CONSTANT
    Terminator : BYTE := 0;
END_VAR
IF NOT EvaluationActive THEN
    RETURN;
END_IF;

IF Result = E_Result.Error THEN
    RETURN;
END_IF;

// C0371: FB inputs are checked before any reference access.
{warning disable C0371}
IF NOT __ISVALIDREF(IN) THEN
    Error(Message := 'Assertion error: IN reference is invalid.');
    RETURN;
END_IF;

IF NOT __ISVALIDREF(Expected) THEN
    Error(Message := 'Assertion error: Expected reference is invalid.');
    RETURN;
END_IF;

IF NOT IsAssertionStringLengthValid(Value := Expected) THEN
    Error(Message := 'Assertion error: Expected exceeds configured STRING length.');
    RETURN;
END_IF;

IF Expected[0] = Terminator THEN
    Error(Message := 'Assertion error: Expected must not be empty.');
    RETURN;
END_IF;

ExpectedLength := 0;
FOR CharacterIndex := 0 TO UINT_TO_DINT(Param_Assertions.AssertionStringLength) DO
    IF Expected[CharacterIndex] = Terminator THEN
        ExpectedLength := CharacterIndex;
        EXIT;
    END_IF;
END_FOR;

InLowerIndex := LOWER_BOUND(IN, 1);
InUpperIndex := UPPER_BOUND(IN, 1);
EndIndex := DINT_TO_LINT(StartIndex) + USINT_TO_LINT(Length) - 1;
IF (Length = 0)
    OR (StartIndex < InLowerIndex) OR (StartIndex > InUpperIndex)
    OR (EndIndex > DINT_TO_LINT(InUpperIndex)) THEN
    Message := CONCAT('Assertion error: array range is invalid. StartIndex = ',
        DINT_TO_STRING(StartIndex));
    Message := CONCAT(Message, ', Length = ');
    Message := CONCAT(Message, USINT_TO_STRING(Length));
    Error(Message := Message);
    RETURN;
END_IF;

IF Result = E_Result.Failed THEN
    RETURN;
END_IF;

PatternFound := FALSE;
IF ExpectedLength = USINT_TO_DINT(Length) THEN
    LastCandidateOffset := 0;
    FOR CandidateOffset := 0 TO LastCandidateOffset DO
        PatternMatches := TRUE;
        FOR CharacterIndex := 0 TO ExpectedLength - 1 DO
            InIndex := LINT_TO_DINT(DINT_TO_LINT(StartIndex) + CandidateOffset
                + DINT_TO_LINT(CharacterIndex));
            IF IN[InIndex] <> Expected[CharacterIndex] THEN
                PatternMatches := FALSE;
                EXIT;
            END_IF;
        END_FOR;
        IF PatternMatches THEN
            PatternFound := TRUE;
            EXIT;
        END_IF;
    END_FOR;
END_IF;

IF NOT PatternFound THEN
    ExpectedText := CreateAssertionTextValue_String(Value := Expected);
    Message := CONCAT('Assertion failed: selected array does not equal Expected = ',
        ExpectedText);
    Message := CONCAT(Message, ', Range = [');
    Message := CONCAT(Message, DINT_TO_STRING(StartIndex));
    Message := CONCAT(Message, '..');
    Message := CONCAT(Message, LINT_TO_STRING(EndIndex));
    Message := CONCAT(Message, '], ExpectedLength = ');
    Message := CONCAT(Message, DINT_TO_STRING(ExpectedLength));
    Message := CONCAT(Message, '.');
    Fail(Message := Message);
    RETURN;
END_IF;

Pass();
{warning restore C0371}
END_METHOD

END_FUNCTION_BLOCK

// ---- Framework/Assertions/POU/Arrays/Char/AssertArrayNoValueChange_Char.TcPOU
{region 'Documentation'}
(*!
<summary>Character codes use BYTE; exact comparison without a mask.</summary>
<description>

Disabling observation preserves the original snapshot. Re-enabling requires a fresh
preceding observation before comparisons resume; it does not replace that snapshot.

StartIndex is an absolute IN index and Length selects 1..255 elements within IN. Memory
must have at least Length elements from its own lower bound. Invalid references or ranges
report Error.

The caller provides dedicated writable Memory that must not overlap IN; overlap is not
checked. Keep bindings, selected range and snapshot contents stable until Reset. Reset
invalidates the snapshot without clearing Memory bytes.

</description>
*)
{endregion}
FUNCTION_BLOCK AssertArrayNoValueChange_Char EXTENDS AssertionBase
VAR_INPUT
    StartIndex : DINT; //! First selected index in IN; uses the array's declared index range, not a zero-based offset.
    Length : USINT; //! Number of monitored elements, from 1 through 255.
END_VAR
VAR_IN_OUT CONSTANT
    IN : ARRAY[*] OF BYTE; //! Read-only actual data; the selected range must remain stable during the call.
END_VAR
VAR_IN_OUT
    Memory : ARRAY[*] OF BYTE; //! Dedicated snapshot storage; only this assertion writes its selected elements.
END_VAR
VAR
    FSnapshotValid : BOOL;
    FObservationPrevious : BOOL;
    FEvaluationActive : BOOL;
END_VAR

SUPER^();

{region 'Documentation'}
(*!
<summary>Capture once or compare against the retained snapshot after range validation.</summary>
*)
{endregion}
METHOD PROTECTED Assert
VAR
    InLowerIndex : DINT;
    InUpperIndex : DINT;
    MemoryLowerIndex : DINT;
    MemoryUpperIndex : DINT;
    MemoryEndIndex : LINT;
    EndIndex : LINT;
    Offset : LINT;
    InIndex : DINT;
    MemoryIndex : DINT;
    Message : STRING(GVL_Constants.MessageLength);
    ReferenceText : STRING;
    ActualText : STRING;
END_VAR
FEvaluationActive := ObservationActive AND FObservationPrevious AND FSnapshotValid;
FObservationPrevious := ObservationActive;

IF NOT ObservationActive THEN
    RETURN;
END_IF;

IF Result = E_Result.Error THEN
    RETURN;
END_IF;

// C0371: FB inputs are checked here before any reference access.
{warning disable C0371}
IF NOT __ISVALIDREF(IN) THEN
    Error(Message := 'Assertion error: IN reference is invalid.');
    RETURN;
END_IF;

IF NOT __ISVALIDREF(Memory) THEN
    Error(Message := 'Assertion error: Memory reference is invalid.');
    RETURN;
END_IF;

InLowerIndex := LOWER_BOUND(IN, 1);
InUpperIndex := UPPER_BOUND(IN, 1);
MemoryLowerIndex := LOWER_BOUND(Memory, 1);
MemoryUpperIndex := UPPER_BOUND(Memory, 1);
EndIndex := DINT_TO_LINT(StartIndex) + USINT_TO_LINT(Length) - 1;
MemoryEndIndex := DINT_TO_LINT(MemoryLowerIndex) + USINT_TO_LINT(Length) - 1;

IF (Length = 0)
    OR (StartIndex < InLowerIndex) OR (StartIndex > InUpperIndex)
    OR (EndIndex > DINT_TO_LINT(InUpperIndex))
    OR (MemoryEndIndex > DINT_TO_LINT(MemoryUpperIndex)) THEN
    Message := CONCAT('Assertion error: array or memory range is invalid. StartIndex = ',
        DINT_TO_STRING(StartIndex));
    Message := CONCAT(Message, ', EndIndex = ');
    Message := CONCAT(Message, LINT_TO_STRING(EndIndex));
    Message := CONCAT(Message, ', Length = ');
    Message := CONCAT(Message, USINT_TO_STRING(Length));
    Message := CONCAT(Message, '.');
    Error(Message := Message);
    RETURN;
END_IF;

IF NOT FSnapshotValid THEN
    FOR Offset := 0 TO USINT_TO_LINT(Length) - 1 DO
        InIndex := LINT_TO_DINT(DINT_TO_LINT(StartIndex) + Offset);
        MemoryIndex := LINT_TO_DINT(DINT_TO_LINT(MemoryLowerIndex) + Offset);
        Memory[MemoryIndex] := IN[InIndex];
    END_FOR;
    FSnapshotValid := TRUE;
    RETURN;
END_IF;

IF NOT EvaluationActive THEN
    RETURN;
END_IF;

IF Result = E_Result.Failed THEN
    RETURN;
END_IF;

FOR Offset := 0 TO USINT_TO_LINT(Length) - 1 DO
    InIndex := LINT_TO_DINT(DINT_TO_LINT(StartIndex) + Offset);
    MemoryIndex := LINT_TO_DINT(DINT_TO_LINT(MemoryLowerIndex) + Offset);
    IF IN[InIndex] <> Memory[MemoryIndex] THEN
        ReferenceText := CreateAssertionTextValue_Char(Value := Memory[MemoryIndex]);
        ActualText := CreateAssertionTextValue_Char(Value := IN[InIndex]);
        Message := CONCAT('Assertion failed: array value changed. Reference[',
            DINT_TO_STRING(MemoryIndex));
        Message := CONCAT(Message, '] = ');
        Message := CONCAT(Message, ReferenceText);
        Message := CONCAT(Message, ', IN[');
        Message := CONCAT(Message, DINT_TO_STRING(InIndex));
        Message := CONCAT(Message, '] = ');
        Message := CONCAT(Message, ActualText);
        Message := CONCAT(Message, '.');
        Fail(Message := Message);
        RETURN;
    END_IF;
END_FOR;

Pass();
{warning restore C0371}
END_METHOD

{region 'Documentation'}
(*!
<summary>Current/last call has consecutive observation and an existing snapshot.</summary>
*)
{endregion}
{attribute 'monitoring' := 'call'}
PROPERTY PUBLIC EvaluationActive : BOOL //! Current/last call has consecutive observation and an existing snapshot.
GET // PUBLIC
EvaluationActive := FEvaluationActive;
END_GET
END_PROPERTY

{region 'Documentation'}
(*!
<summary>Invalidate the snapshot and observation history.</summary>
<description>

Does not clear external Memory. The next active observation captures a new snapshot
before comparison.

</description>
*)
{endregion}
METHOD PROTECTED ResetAssertion
FSnapshotValid := FALSE;
FObservationPrevious := FALSE;
FEvaluationActive := FALSE;
END_METHOD

END_FUNCTION_BLOCK

// ---- Framework/Assertions/POU/Arrays/Char/AssertArrayStartsWithString_Char.TcPOU
{region 'Documentation'}
(*!
<summary>Check that the selected array starts with the STRING code units.</summary>
<description>

StartIndex is an absolute declared IN index, not an offset. Length selects 1..255
elements; the complete selected range must fit IN. Invalid references or ranges report
Error.

Keep supplied arrays stable for the call. Input data is read, not copied or retained as a
snapshot.

Expected must be nonempty and fit its configured text capacity (otherwise Error). A valid
text longer than the selected array region reports Failed. The array is not zero-terminated or
trimmed; matching is exact and case-sensitive.

</description>
*)
{endregion}
FUNCTION_BLOCK AssertArrayStartsWithString_Char EXTENDS AssertionBase
VAR_INPUT
    StartIndex : DINT; //! First selected index in IN; uses the array's declared index range, not a zero-based offset.
    Length : USINT; //! Number of selected array elements, from 1 through 255.
END_VAR
VAR_IN_OUT CONSTANT
    IN : ARRAY[*] OF BYTE; //! Read-only actual data; the selected range must remain stable during the call.
    Expected : STRING(Param_Assertions.AssertionStringLength); //! Nonempty expected text, terminated within the configured capacity; keep stable during the call.
END_VAR

SUPER^();

{region 'Documentation'}
(*!
<summary>Validate references and ranges before exact code-unit comparison.</summary>
*)
{endregion}
METHOD PROTECTED Assert
VAR
    InLowerIndex : DINT;
    InUpperIndex : DINT;
    EndIndex : LINT;
    ExpectedLength : DINT;
    CharacterIndex : DINT;
    InIndex : DINT;
    CandidateOffset : LINT;
    LastCandidateOffset : LINT;
    PatternMatches : BOOL;
    PatternFound : BOOL;
    ExpectedText : STRING(GVL_Constants.AssertionValueLength);
    Message : STRING(GVL_Constants.MessageLength);
END_VAR
VAR CONSTANT
    Terminator : BYTE := 0;
END_VAR
IF NOT EvaluationActive THEN
    RETURN;
END_IF;

IF Result = E_Result.Error THEN
    RETURN;
END_IF;

// C0371: FB inputs are checked before any reference access.
{warning disable C0371}
IF NOT __ISVALIDREF(IN) THEN
    Error(Message := 'Assertion error: IN reference is invalid.');
    RETURN;
END_IF;

IF NOT __ISVALIDREF(Expected) THEN
    Error(Message := 'Assertion error: Expected reference is invalid.');
    RETURN;
END_IF;

IF NOT IsAssertionStringLengthValid(Value := Expected) THEN
    Error(Message := 'Assertion error: Expected exceeds configured STRING length.');
    RETURN;
END_IF;

IF Expected[0] = Terminator THEN
    Error(Message := 'Assertion error: Expected must not be empty.');
    RETURN;
END_IF;

ExpectedLength := 0;
FOR CharacterIndex := 0 TO UINT_TO_DINT(Param_Assertions.AssertionStringLength) DO
    IF Expected[CharacterIndex] = Terminator THEN
        ExpectedLength := CharacterIndex;
        EXIT;
    END_IF;
END_FOR;

InLowerIndex := LOWER_BOUND(IN, 1);
InUpperIndex := UPPER_BOUND(IN, 1);
EndIndex := DINT_TO_LINT(StartIndex) + USINT_TO_LINT(Length) - 1;
IF (Length = 0)
    OR (StartIndex < InLowerIndex) OR (StartIndex > InUpperIndex)
    OR (EndIndex > DINT_TO_LINT(InUpperIndex)) THEN
    Message := CONCAT('Assertion error: array range is invalid. StartIndex = ',
        DINT_TO_STRING(StartIndex));
    Message := CONCAT(Message, ', Length = ');
    Message := CONCAT(Message, USINT_TO_STRING(Length));
    Error(Message := Message);
    RETURN;
END_IF;

IF Result = E_Result.Failed THEN
    RETURN;
END_IF;

PatternFound := FALSE;
IF ExpectedLength <= USINT_TO_DINT(Length) THEN
    LastCandidateOffset := 0;
    FOR CandidateOffset := 0 TO LastCandidateOffset DO
        PatternMatches := TRUE;
        FOR CharacterIndex := 0 TO ExpectedLength - 1 DO
            InIndex := LINT_TO_DINT(DINT_TO_LINT(StartIndex) + CandidateOffset
                + DINT_TO_LINT(CharacterIndex));
            IF IN[InIndex] <> Expected[CharacterIndex] THEN
                PatternMatches := FALSE;
                EXIT;
            END_IF;
        END_FOR;
        IF PatternMatches THEN
            PatternFound := TRUE;
            EXIT;
        END_IF;
    END_FOR;
END_IF;

IF NOT PatternFound THEN
    ExpectedText := CreateAssertionTextValue_String(Value := Expected);
    Message := CONCAT('Assertion failed: selected array does not start with Expected = ',
        ExpectedText);
    Message := CONCAT(Message, ', Range = [');
    Message := CONCAT(Message, DINT_TO_STRING(StartIndex));
    Message := CONCAT(Message, '..');
    Message := CONCAT(Message, LINT_TO_STRING(EndIndex));
    Message := CONCAT(Message, '], ExpectedLength = ');
    Message := CONCAT(Message, DINT_TO_STRING(ExpectedLength));
    Message := CONCAT(Message, '.');
    Fail(Message := Message);
    RETURN;
END_IF;

Pass();
{warning restore C0371}
END_METHOD

END_FUNCTION_BLOCK

// ---- Framework/Assertions/POU/Arrays/Char/AssertEqualArray_Char.TcPOU
{region 'Documentation'}
(*!
<summary>Character codes use BYTE; exact comparison without a mask.</summary>
<description>

Compares the entire Expected array with IN starting at StartIndex.

StartIndex is an absolute declared IN index. The entire Expected array, starting at its
own lower bound, determines the compared length and must fit IN. Invalid references or ranges
report Error.

Keep supplied arrays stable for the call. Input data is read, not copied or retained as a
snapshot.

</description>
*)
{endregion}
FUNCTION_BLOCK AssertEqualArray_Char EXTENDS AssertionBase
VAR_INPUT
    StartIndex : DINT; //! First compared index in IN; Expected starts at its own lower bound.
END_VAR
VAR_IN_OUT CONSTANT
    IN : ARRAY[*] OF BYTE; //! Read-only actual data; the selected range must remain stable during the call.
    Expected : ARRAY[*] OF BYTE; //! Read-only expected sequence starting at its own lower bound; must fit the selected actual range.
END_VAR

SUPER^();

{region 'Documentation'}
(*!
<summary>Validate the selected range and expectations before comparing elements.</summary>
*)
{endregion}
METHOD PROTECTED Assert
VAR
    InLowerIndex : DINT;
    InUpperIndex : DINT;
    ExpectedLowerIndex : DINT;
    ExpectedUpperIndex : DINT;
    ExpectedLength : LINT;
    EndIndex : LINT;
    Offset : LINT;
    InIndex : DINT;
    ExpectedIndex : DINT;
    Message : STRING(GVL_Constants.MessageLength);
    ExpectedText : STRING;
    ActualText : STRING;
END_VAR
IF NOT EvaluationActive THEN
    RETURN;
END_IF;

IF Result = E_Result.Error THEN
    RETURN;
END_IF;

// C0371: FB inputs are checked here before any reference access.
{warning disable C0371}
IF NOT __ISVALIDREF(IN) THEN
    Error(Message := 'Assertion error: IN reference is invalid.');
    RETURN;
END_IF;

IF NOT __ISVALIDREF(Expected) THEN
    Error(Message := 'Assertion error: Expected reference is invalid.');
    RETURN;
END_IF;

InLowerIndex := LOWER_BOUND(IN, 1);
InUpperIndex := UPPER_BOUND(IN, 1);
ExpectedLowerIndex := LOWER_BOUND(Expected, 1);
ExpectedUpperIndex := UPPER_BOUND(Expected, 1);
ExpectedLength := DINT_TO_LINT(ExpectedUpperIndex) - DINT_TO_LINT(ExpectedLowerIndex) + 1;
EndIndex := DINT_TO_LINT(StartIndex) + ExpectedLength - 1;

